// TwinCAT 3 PLC project test
// ProgramVersion: 3.1.4026.27
// libraries:
//   Tc2_Standard, * (Beckhoff Automation GmbH)
//   Tc2_System, * (Beckhoff Automation GmbH)
//   Tc2_Utilities, * (Beckhoff Automation GmbH)
//   Tc3_IotBase, * (Beckhoff Automation GmbH)
//   Tc3_JsonXml, * (Beckhoff Automation GmbH)
//   TcOtlp, * (S&E Engineering)
//   TcUnit, * (www.tcunit.org)
// project tree:
//   / MAIN.TcPOU, PlcTask.TcTTO
//   TEST/TRACING/EXPORTING/ FB_SpanExporter_ForInspection.TcPOU, FB_TestSpanFileExporter.TcPOU, FB_TestSpanSimulation.TcPOU, FB_TestSpanConsoleExporter.TcPOU, FB_TestSpanHttpExporter.TcPOU
//   TEST/EXPORTING/ FB_TestHttpUrlParser.TcPOU
//   TEST/TRACING/TRACESTATE/ FB_TestTraceState.TcPOU
//   TEST/TRACING/PROPAGATION/ FB_TestTraceContextPropagator.TcPOU, FB_TestAdsLoopbackPropagation.TcPOU
//   TEST/TRACING/SAMPLING/ FB_Sampler_ForInspection.TcPOU, FB_TestSamplers.TcPOU
//   TEST/LOGGING/EXPORTING/ FB_TestFileExporter.TcPOU, FB_TestHttpExporter.TcPOU, FB_TestLogExporters.TcPOU
//   TEST/LOGGING/EXPORTING/UTILS/ FB_LogRecordExporter_File_ForSerializationInspection.TcPOU, FB_LogRecordExporter_ForInspection.TcPOU
//   TEST/LOGGING/LOGGER/ FB_TestLogger.TcPOU
//   TEST/LOGGING/LOG_RECORD/ FB_TestLogRecord.TcPOU, FB_TestLogRecordQueue.TcPOU
//   TEST/LOGGING/PROCESSOR/ FB_TestLogProcessors.TcPOU
//   TEST/LOGGING/PROCESSOR/UTILS/ FB_LogRecordProcessor_ConsolePrinter.TcPOU, FB_LogRecordProcessor_ForBatchInspection.TcPOU, FB_LogRecordProcessor_ForRecordInspection.TcPOU, FB_LogRecordProcessor_ForRecordsInspection.TcPOU
//   TEST/LOGGING/PROVIDER/ FB_TestLoggerProvider.TcPOU
//   TEST/LOGGING/SERIALIZATION/ FB_TestProtoJsonSerializer.TcPOU
//   TEST/TRACING/ID_GENERATOR/ FB_TestIdGenerator.TcPOU
//   TEST/TRACING/PROCESSOR/ FB_SpanProcessor_ForInspection.TcPOU, FB_TestSpanProcessors.TcPOU
//   TEST/TRACING/PROVIDER/ FB_TestTracerProvider.TcPOU, FB_TracerProvider_ForInspection.TcPOU
//   TEST/TRACING/TRACER/ FB_MockIdGenerator.TcPOU, FB_TestTracer.TcPOU
//   TEST/TRACING/LINK/ FB_TestLinks.TcPOU
//   TEST/TRACING/SERIALIZATION/ FB_TestSpanProtoJsonSerializer.TcPOU
//   TEST/TRACING/SPAN/ FB_TestSpan.TcPOU, FB_TestSpanContext.TcPOU, FB_TestSpanQueue.TcPOU
//   TEST/VALUES/ FB_TestAttributes.TcPOU, FB_TestOtlpValue.TcPOU
// real-time tasks:
//   TASK PlcTask: cycle T#10ms, priority 20, ADS port 350

CONFIGURATION test
    RESOURCE PLC ON TwinCAT3
        TASK PlcTask(INTERVAL := T#10ms, PRIORITY := 20);
        PROGRAM MAIN WITH PlcTask : MAIN;
    END_RESOURCE
END_CONFIGURATION

// ---- MAIN.TcPOU
PROGRAM MAIN
VAR
	{attribute 'analysis' := '-33'}fbTestOtlpValue: FB_TestOtlpValue();
	{attribute 'analysis' := '-33'}fbTestAttributes: FB_TestAttributes();
	{attribute 'analysis' := '-33'}fbTestLogRecordQueue: FB_TestLogRecordQueue();
	{attribute 'analysis' := '-33'}fbTestLogger: FB_TestLogger();
	{attribute 'analysis' := '-33'}fbTestProvider: FB_TestLoggerProvider();
	{attribute 'analysis' := '-33'}fbTestProcessors: FB_TestLogProcessors();
	{attribute 'analysis' := '-33'}fbTestExporters: FB_TestLogExporters();
	{attribute 'analysis' := '-33'}fbTestLogRecord: FB_TestLogRecord();
	{attribute 'analysis' := '-33'}fbTestProtoJsonSerializer: FB_TestProtoJsonSerializer();
	{attribute 'analysis' := '-33'}fbTestFileExporter: FB_TestFileExporter();
	{attribute 'analysis' := '-33'}fbTestHttpExporter: FB_TestHttpExporter();
	{attribute 'analysis' := '-33'}fbTestIdGenerator: FB_TestIdGenerator();
	{attribute 'analysis' := '-33'}fbTestSpanContext: FB_TestSpanContext();
	{attribute 'analysis' := '-33'}fbTestTraceState: FB_TestTraceState();
	{attribute 'analysis' := '-33'}fbTestTraceContextPropagator: FB_TestTraceContextPropagator();
	{attribute 'analysis' := '-33'}fbTestAdsLoopbackPropagation: FB_TestAdsLoopbackPropagation();
	{attribute 'analysis' := '-33'}fbTestSpan: FB_TestSpan();
	{attribute 'analysis' := '-33'}fbTestTracer: FB_TestTracer();
	{attribute 'analysis' := '-33'}fbTestSpanQueue: FB_TestSpanQueue();
	{attribute 'analysis' := '-33'}fbTestSpanProcessors: FB_TestSpanProcessors();
	{attribute 'analysis' := '-33'}fbTestTracerProvider: FB_TestTracerProvider();
	{attribute 'analysis' := '-33'}fbTestSamplers: FB_TestSamplers();
	{attribute 'analysis' := '-33'}fbTestSpanProtoJsonSerializer: FB_TestSpanProtoJsonSerializer();
	{attribute 'analysis' := '-33'}fbTestLinks: FB_TestLinks();
	{attribute 'analysis' := '-33'}fbTestSpanFileExporter: FB_TestSpanFileExporter();
	{attribute 'analysis' := '-33'}fbTestSpanConsoleExporter: FB_TestSpanConsoleExporter();
	{attribute 'analysis' := '-33'}fbTestSpanHttpExporter: FB_TestSpanHttpExporter();
	{attribute 'analysis' := '-33'}fbTestHttpUrlParser: FB_TestHttpUrlParser();
	{attribute 'analysis' := '-33'}fbTestSpanSimulation: FB_TestSpanSimulation();
END_VAR

TcUnit.RUN();

END_PROGRAM

// ---- TEST/VALUES/FB_TestOtlpValue.TcPOU
(* Tests that ValueFactory validates its inputs, copies what it is given, and that every value it builds is released exactly once. *)
FUNCTION_BLOCK FB_TestOtlpValue EXTENDS FB_TestSuite

THIS^.testCreateStringValidatesInputs();
THIS^.testCreateTraceIdCopiesBytes();
THIS^.testCreateSpanIdCopiesBytes();
THIS^.testCreateKeyValueValidatesInputs();
THIS^.testCreateNumberCopiesEveryNumericType();
THIS^.testCloneCopiesAndForwardsFailures();
THIS^.testDeleteClearsPointer();

(* delete releases a value and clears the caller's pointer, through the concrete or the base type, and refuses a pointer to another value so nothing is released twice. *)
METHOD testDeleteClearsPointer : REFERENCE TO FB_Test
VAR
	pStr: POINTER TO FB_String;
	pOther: POINTER TO FB_String;
	pAny: POINTER TO FB_AnyValue;
	pOtherBefore: POINTER TO FB_String;
	deleted: BOOL;
	failureReason: E_ValueFactoryFailureReason;
END_VAR
TcUnit.TEST('testDeleteClearsPointer');

	// through the concrete pointer type
	IF ValueFactory.createString(pDest:=pStr, pString:=ADR('value'), failureReason=>failureReason) THEN
		deleted := pStr^.delete(pSelf:=pStr);
		THIS^.AssertTrue(deleted, 'Expected delete through an FB_String pointer to succeed');
		THIS^.AssertTrue(pStr = 0, 'Expected delete to clear the FB_String pointer');
	ELSE
		THIS^.AssertTrue(FALSE, 'Expected createString to succeed for the FB_String pointer case');
	END_IF

	// through the abstract base pointer, dispatched to FB_String
	IF ValueFactory.createString(pDest:=pStr, pString:=ADR('value'), failureReason=>failureReason) THEN
		pAny := pStr;
		pStr := 0;
		deleted := pAny^.delete(pSelf:=pAny);
		THIS^.AssertTrue(deleted, 'Expected delete through an FB_AnyValue pointer to succeed');
		THIS^.AssertTrue(pAny = 0, 'Expected delete to clear the FB_AnyValue pointer');
	ELSE
		THIS^.AssertTrue(FALSE, 'Expected createString to succeed for the FB_AnyValue pointer case');
	END_IF

	// a pointer to another value is refused and left untouched
	IF ValueFactory.createString(pDest:=pStr, pString:=ADR('first'), failureReason=>failureReason)
		AND_THEN ValueFactory.createString(pDest:=pOther, pString:=ADR('second'), failureReason=>failureReason)
	THEN
		pOtherBefore := pOther;
		deleted := pStr^.delete(pSelf:=pOther);
		THIS^.AssertFalse(deleted, 'Expected delete with another value$'s pointer to be refused');
		THIS^.AssertTrue(pOther = pOtherBefore, 'Expected a refused delete to leave the pointer unchanged');
		THIS^.AssertEquals_STRING(Expected:='first', Actual:=pStr^.pString^, Message:='Expected the first value to survive a refused delete');
		THIS^.AssertEquals_STRING(Expected:='second', Actual:=pOther^.pString^, Message:='Expected the second value to survive a refused delete');
	ELSE
		THIS^.AssertTrue(FALSE, 'Expected createString to succeed for both strings of the refused delete case');
	END_IF
	IF pStr <> 0 THEN pStr^.delete(pSelf:=pStr); END_IF
	IF pOther <> 0 THEN pOther^.delete(pSelf:=pOther); END_IF

TcUnit.TEST_FINISHED();
END_METHOD

(*
	The clone functions copy strings, numbers, and key values into new allocations.
	A nested clone failure is forwarded with its reason and leaves the destination unassigned, so a caller never gets a half-built value.
*)
METHOD testCloneCopiesAndForwardsFailures : REFERENCE TO FB_Test
VAR
	pStringSource: POINTER TO FB_String;
	pStringClone: POINTER TO FB_String;
	pNumberSource: POINTER TO FB_Number;
	pNumberClone: POINTER TO FB_Number;
	pKeyValueSource: POINTER TO FB_KeyValue;
	pKeyValueClone: POINTER TO FB_KeyValue;
	pAnySource: POINTER TO FB_AnyValue;
	pAnyClone: POINTER TO FB_AnyValue;
	number: DINT := 42;
	success: BOOL;
	failureReason: E_ValueFactoryFailureReason;
	noFailure: E_ValueFactoryFailureReason;
END_VAR
TcUnit.TEST('testCloneCopiesAndForwardsFailures');

	noFailure := E_ValueFactoryFailureReason.NA;

	// cloneString
	success := ValueFactory.createString(pDest:=pStringSource, pString:=ADR('source'), failureReason=>failureReason);
	THIS^.AssertTrue(success AND_THEN failureReason=noFailure AND_THEN pStringSource<>0, 'Expected createString to build the source string');

	success := ValueFactory.cloneString(pDest:=pStringClone, pSrc:=pStringSource, failureReason=>failureReason);
	THIS^.AssertTrue(success AND_THEN failureReason=noFailure AND_THEN pStringClone<>0, 'Expected cloneString to succeed');
	IF pStringClone <> 0 THEN
		THIS^.AssertEquals_STRING('source', pStringClone^.pString^, 'Expected cloneString to copy the source text');
		pStringClone^.delete(pSelf:=pStringClone);
	END_IF

	// cloneNumber
	success := ValueFactory.createNumber(pDest:=pNumberSource, value:=number, failureReason=>failureReason);
	THIS^.AssertTrue(success AND_THEN failureReason=noFailure AND_THEN pNumberSource<>0, 'Expected createNumber to build the source number');

	success := ValueFactory.cloneNumber(pDest:=pNumberClone, pSrc:=pNumberSource, failureReason=>failureReason);
	THIS^.AssertTrue(success AND_THEN failureReason=noFailure AND_THEN pNumberClone<>0, 'Expected cloneNumber to succeed');
	IF pNumberClone <> 0 THEN
		THIS^.AssertTrue(MEMCMP(pNumberClone^.value.pValue, ADR(number), SIZEOF(number))=0, 'Expected cloneNumber to copy the source value');
		pNumberClone^.delete(pSelf:=pNumberClone);
	END_IF

	// cloneAnyValue dispatches on the value type
	pAnySource := pNumberSource;
	success := ValueFactory.cloneAnyValue(pDest:=pAnyClone, pSrc:=pAnySource, failureReason=>failureReason);
	THIS^.AssertTrue(success AND_THEN failureReason=noFailure AND_THEN pAnyClone<>0, 'Expected cloneAnyValue to forward a successful number clone');
	IF pAnyClone <> 0 THEN
		THIS^.AssertTrue(pAnyClone^.eType=E_ValueType.E_Number, 'Expected cloneAnyValue to produce a number');
		pAnyClone^.delete(pSelf:=pAnyClone);
	END_IF

	// cloneKeyValue
	success := ValueFactory.createKeyValue(pDest:=pKeyValueSource, pKey:=ADR('key'), pVal:=pStringSource, failureReason=>failureReason);
	THIS^.AssertTrue(success AND_THEN failureReason=noFailure AND_THEN pKeyValueSource<>0, 'Expected createKeyValue to build the source key value');

	success := ValueFactory.cloneKeyValue(pDest:=pKeyValueClone, pSrc:=pKeyValueSource, failureReason=>failureReason);
	THIS^.AssertTrue(success AND_THEN failureReason=noFailure AND_THEN pKeyValueClone<>0, 'Expected cloneKeyValue to succeed');
	IF pKeyValueClone <> 0 THEN
		THIS^.AssertEquals_STRING('key', pKeyValueClone^.pKey^, 'Expected cloneKeyValue to copy the source key');
		pKeyValueClone^.delete(pSelf:=pKeyValueClone);
	END_IF

	// cloneAnyValue must forward a nested cloneString failure without assigning the destination.
	// free() empties the source string, a state the factory would never build, so the nested clone fails.
	IF pStringSource <> 0 THEN pStringSource^.free(); END_IF
	pAnySource := pStringSource;
	success := ValueFactory.cloneAnyValue(pDest:=pAnyClone, pSrc:=pAnySource, failureReason=>failureReason);
	THIS^.AssertFalse(success, 'Expected cloneAnyValue to reject a string with a null payload');
	THIS^.AssertTrue(failureReason=E_ValueFactoryFailureReason.STRING_POINTER_NULL, 'Expected cloneAnyValue to forward the cloneString failure reason');
	THIS^.AssertTrue(pAnyClone=0, 'Expected a failed cloneAnyValue to leave the destination unassigned');

	// cloneKeyValue must forward the nested createKeyValue failure reason.
	// free() empties the source key value, so it has no key to clone.
	IF pKeyValueSource <> 0 THEN pKeyValueSource^.free(); END_IF
	success := ValueFactory.cloneKeyValue(pDest:=pKeyValueClone, pSrc:=pKeyValueSource, failureReason=>failureReason);
	THIS^.AssertFalse(success, 'Expected cloneKeyValue to reject a key value with a null key');
	THIS^.AssertTrue(failureReason=E_ValueFactoryFailureReason.KEY_POINTER_NULL, 'Expected cloneKeyValue to forward the createKeyValue failure reason');
	THIS^.AssertTrue(pKeyValueClone=0, 'Expected a failed cloneKeyValue to leave the destination unassigned');

	IF pStringSource <> 0 THEN pStringSource^.delete(pSelf:=pStringSource); END_IF
	IF pNumberSource <> 0 THEN pNumberSource^.delete(pSelf:=pNumberSource); END_IF
	IF pKeyValueSource <> 0 THEN pKeyValueSource^.delete(pSelf:=pKeyValueSource); END_IF

TcUnit.TEST_FINISHED();
END_METHOD

(*
	createKeyValue rejects a null key, a null value, or an assigned destination with a distinct reason and allocates nothing.
	On success the key value owns its own copy of the value, so the caller may delete the original.
*)
METHOD testCreateKeyValueValidatesInputs : REFERENCE TO FB_Test
VAR
	pKeyVal: POINTER TO FB_KeyValue;
	pVal: POINTER TO FB_String;
	anyValue: POINTER TO FB_AnyValue;
	expectedType: E_ValueType := E_ValueType.E_KeyValue;
	actualType: E_ValueType;
	pOriginal: POINTER TO FB_KeyValue;
	success: BOOL;
	failureReason: E_ValueFactoryFailureReason;
	noFailure: E_ValueFactoryFailureReason;
	failureCode: INT;
END_VAR
TcUnit.TEST('testCreateKeyValueValidatesInputs');
	noFailure := E_ValueFactoryFailureReason.NA;

	// null key and null value are rejected
	success := ValueFactory.createKeyValue(pDest:=pKeyVal, pKey:=0, pVal:=0, failureReason=>failureReason);
	THIS^.AssertFalse(success, 'Expected createKeyValue to reject a null key pointer');
	THIS^.AssertTrue(failureReason=E_ValueFactoryFailureReason.KEY_POINTER_NULL, 'Expected the null key failure reason');
	THIS^.AssertTrue(pKeyVal=0, 'Expected a null key to leave the destination unassigned');

	success := ValueFactory.createKeyValue(pDest:=pKeyVal, pKey:=ADR('Key'), pVal:=0, failureReason=>failureReason);
	THIS^.AssertFalse(success, 'Expected createKeyValue to reject a null value pointer');
	THIS^.AssertTrue(failureReason=E_ValueFactoryFailureReason.VALUE_POINTER_NULL, 'Expected the null value failure reason');
	THIS^.AssertTrue(pKeyVal=0, 'Expected a null value to leave the destination unassigned');

	// a valid key and value
	success := ValueFactory.createString(pDest:=pVal, pString:=ADR('Value'), failureReason=>failureReason);
	THIS^.AssertTrue(success AND_THEN failureReason=noFailure AND_THEN pVal<>0, 'Expected createString to build the source value');
	success := ValueFactory.createKeyValue(pDest:=pKeyVal, pKey:=ADR('Key'), pVal:=pVal, failureReason=>failureReason);
	THIS^.AssertTrue(success, 'Expected createKeyValue to succeed with a valid key and value');
	THIS^.AssertTrue(failureReason=noFailure, 'Expected a successful createKeyValue to clear the failure reason');
	THIS^.AssertTrue(pKeyVal<>0, 'Expected a successful createKeyValue to allocate the destination');

	// an assigned destination is refused and left as it was
	pOriginal := pKeyVal;
	success := ValueFactory.createKeyValue(pDest:=pKeyVal, pKey:=ADR('Key'), pVal:=pVal, failureReason=>failureReason);
	THIS^.AssertFalse(success, 'Expected createKeyValue to reject an assigned destination');
	THIS^.AssertTrue(failureReason=E_ValueFactoryFailureReason.DESTINATION_ALREADY_ASSIGNED, 'Expected the assigned destination failure reason');
	THIS^.AssertTrue(pKeyVal=pOriginal, 'Expected a refused createKeyValue to keep the existing destination');
	// E_ValueFactoryFailureReason is numbered implicitly after NA := 0; this pins the first failure code at 1
	// so the numeric codes seen in logs and on an HMI do not shift if the enum declaration is edited.
	failureCode := E_ValueFactoryFailureReason.DESTINATION_ALREADY_ASSIGNED;
	THIS^.AssertEquals_INT(1, failureCode, 'Expected the first ValueFactory failure code to be 1');

 	IF pVal <> 0 AND pKeyVal <> 0 THEN
		// a key value is an FB_AnyValue of type E_KeyValue
		anyValue := pKeyVal;
		actualType := anyValue^.eType;
		THIS^.AssertEquals(
			expectedType,
			actualType,
			'Expected the key value to report the E_KeyValue type'
		);
		THIS^.AssertEquals_STRING(
			Actual:=pKeyVal^.pKey^,
			Expected:='Key',
			Message:='Expected the key value to hold the key'
		);
		// deleting the caller's value proves the key value holds its own copy
		pVal^.delete(pSelf:=pVal);
		pVal := pKeyVal^.pVal;
		THIS^.AssertEquals_STRING(
			Actual:=pVal^.pString^,
			Expected:='Value',
			Message:='Expected the key value to keep its value after the original is deleted'
		);
	END_IF
	// cleanup data
	IF pKeyVal <> 0 THEN pKeyVal^.delete(pSelf:=pKeyVal);
	ELSIF pVal <> 0 THEN pVal^.delete(pSelf:=pVal); END_IF


TcUnit.TEST_FINISHED();
END_METHOD

(*
	createNumber accepts every IEC numeric type and keeps its type class and its own copy of the bytes, so the serializer can write the exact type the caller used.
	It also refuses an assigned destination, and free releases the owned data.
*)
METHOD testCreateNumberCopiesEveryNumericType : REFERENCE TO FB_Test
VAR
	nSInt: SINT := -12;
	nInt: INT := -1234;
	nDInt: DINT := -12345;
	nLInt: LINT := -123456;
	nUSInt: USINT := 12;
	nUInt: UINT := 1234;
	nUDInt: UDINT := 12345;
	nULInt: ULINT := 123456;
	fReal: REAL := 42.25;
	fLReal: LREAL := 24.5;
	pValue: POINTER TO FB_Number;
	pDInt: POINTER TO DINT;
	pOriginal: POINTER TO FB_Number;
	anyValue: POINTER TO FB_AnyValue;
	success: BOOL;
	failureReason: E_ValueFactoryFailureReason;
	noFailure: E_ValueFactoryFailureReason;
END_VAR
TcUnit.TEST('testCreateNumberCopiesEveryNumericType');
noFailure := E_ValueFactoryFailureReason.NA;

// ANY_NUM accepts every signed, unsigned, and floating-point IEC numeric type.

// SINT
success := ValueFactory.createNumber(pDest:=pValue, value:=nSInt, failureReason=>failureReason);
THIS^.AssertTrue(success AND_THEN failureReason=noFailure AND_THEN pValue<>0, 'Expected createNumber to accept a SINT');
IF pValue <> 0 THEN
	THIS^.AssertTrue(pValue^.value.typeclass=__SYSTEM.TYPE_CLASS.TYPE_SINT, 'Expected the SINT type to be kept');
	THIS^.AssertTrue(pValue^.value.diSize=SIZEOF(nSInt) AND_THEN MEMCMP(pValue^.value.pValue, ADR(nSInt), SIZEOF(nSInt))=0, 'Expected the SINT value to be copied');
	pValue^.delete(pSelf:=pValue);
END_IF

// INT
success := ValueFactory.createNumber(pDest:=pValue, value:=nInt, failureReason=>failureReason);
THIS^.AssertTrue(success AND_THEN failureReason=noFailure AND_THEN pValue<>0, 'Expected createNumber to accept an INT');
IF pValue <> 0 THEN
	THIS^.AssertTrue(pValue^.value.typeclass=__SYSTEM.TYPE_CLASS.TYPE_INT, 'Expected the INT type to be kept');
	THIS^.AssertTrue(pValue^.value.diSize=SIZEOF(nInt) AND_THEN MEMCMP(pValue^.value.pValue, ADR(nInt), SIZEOF(nInt))=0, 'Expected the INT value to be copied');
	pValue^.delete(pSelf:=pValue);
END_IF

// DINT, plus copy independence and an assigned destination
success := ValueFactory.createNumber(pDest:=pValue, value:=nDInt, failureReason=>failureReason);
THIS^.AssertTrue(success AND_THEN failureReason=noFailure AND_THEN pValue<>0, 'Expected createNumber to accept a DINT');
IF pValue <> 0 THEN
	THIS^.AssertTrue(pValue^.value.typeclass=__SYSTEM.TYPE_CLASS.TYPE_DINT, 'Expected the DINT type to be kept');
	THIS^.AssertTrue(pValue^.value.diSize=SIZEOF(nDInt) AND_THEN MEMCMP(pValue^.value.pValue, ADR(nDInt), SIZEOF(nDInt))=0, 'Expected the DINT value to be copied');
	// The wrapper owns a copy; changing the source must not change the wrapped value.
	pDInt := pValue^.value.pValue;
	nDInt := 7;
	THIS^.AssertEquals_DINT(-12345, pDInt^, 'Expected the number to keep its value after the source DINT changes');
	// A factory call must never replace an already allocated destination.
	pOriginal := pValue;
	success := ValueFactory.createNumber(pDest:=pValue, value:=fLReal, failureReason=>failureReason);
	THIS^.AssertFalse(success, 'Expected createNumber to reject an allocated destination');
	THIS^.AssertTrue(failureReason=E_ValueFactoryFailureReason.DESTINATION_ALREADY_ASSIGNED, 'Expected the assigned number destination failure reason');
	THIS^.AssertTrue(pValue=pOriginal, 'Expected a refused createNumber to keep the existing destination');
	pValue^.delete(pSelf:=pValue);
END_IF

// LINT, which also proves the previous failure reason is cleared
success := ValueFactory.createNumber(pDest:=pValue, value:=nLInt, failureReason=>failureReason);
THIS^.AssertTrue(success AND_THEN failureReason=noFailure AND_THEN pValue<>0, 'Expected createNumber to accept a LINT and clear the previous failure reason');
IF pValue <> 0 THEN
	THIS^.AssertTrue(pValue^.value.typeclass=__SYSTEM.TYPE_CLASS.TYPE_LINT, 'Expected the LINT type to be kept');
	THIS^.AssertTrue(pValue^.value.diSize=SIZEOF(nLInt) AND_THEN MEMCMP(pValue^.value.pValue, ADR(nLInt), SIZEOF(nLInt))=0, 'Expected the LINT value to be copied');
	pValue^.delete(pSelf:=pValue);
END_IF

// USINT
success := ValueFactory.createNumber(pDest:=pValue, value:=nUSInt, failureReason=>failureReason);
THIS^.AssertTrue(success AND_THEN failureReason=noFailure AND_THEN pValue<>0, 'Expected createNumber to accept a USINT');
IF pValue <> 0 THEN
	THIS^.AssertTrue(pValue^.value.typeclass=__SYSTEM.TYPE_CLASS.TYPE_USINT, 'Expected the USINT type to be kept');
	THIS^.AssertTrue(pValue^.value.diSize=SIZEOF(nUSInt) AND_THEN MEMCMP(pValue^.value.pValue, ADR(nUSInt), SIZEOF(nUSInt))=0, 'Expected the USINT value to be copied');
	pValue^.delete(pSelf:=pValue);
END_IF

// UINT
success := ValueFactory.createNumber(pDest:=pValue, value:=nUInt, failureReason=>failureReason);
THIS^.AssertTrue(success AND_THEN failureReason=noFailure AND_THEN pValue<>0, 'Expected createNumber to accept a UINT');
IF pValue <> 0 THEN
	THIS^.AssertTrue(pValue^.value.typeclass=__SYSTEM.TYPE_CLASS.TYPE_UINT, 'Expected the UINT type to be kept');
	THIS^.AssertTrue(pValue^.value.diSize=SIZEOF(nUInt) AND_THEN MEMCMP(pValue^.value.pValue, ADR(nUInt), SIZEOF(nUInt))=0, 'Expected the UINT value to be copied');
	pValue^.delete(pSelf:=pValue);
END_IF

// UDINT
success := ValueFactory.createNumber(pDest:=pValue, value:=nUDInt, failureReason=>failureReason);
THIS^.AssertTrue(success AND_THEN failureReason=noFailure AND_THEN pValue<>0, 'Expected createNumber to accept a UDINT');
IF pValue <> 0 THEN
	THIS^.AssertTrue(pValue^.value.typeclass=__SYSTEM.TYPE_CLASS.TYPE_UDINT, 'Expected the UDINT type to be kept');
	THIS^.AssertTrue(pValue^.value.diSize=SIZEOF(nUDInt) AND_THEN MEMCMP(pValue^.value.pValue, ADR(nUDInt), SIZEOF(nUDInt))=0, 'Expected the UDINT value to be copied');
	pValue^.delete(pSelf:=pValue);
END_IF

// ULINT
success := ValueFactory.createNumber(pDest:=pValue, value:=nULInt, failureReason=>failureReason);
THIS^.AssertTrue(success AND_THEN failureReason=noFailure AND_THEN pValue<>0, 'Expected createNumber to accept a ULINT');
IF pValue <> 0 THEN
	THIS^.AssertTrue(pValue^.value.typeclass=__SYSTEM.TYPE_CLASS.TYPE_ULINT, 'Expected the ULINT type to be kept');
	THIS^.AssertTrue(pValue^.value.diSize=SIZEOF(nULInt) AND_THEN MEMCMP(pValue^.value.pValue, ADR(nULInt), SIZEOF(nULInt))=0, 'Expected the ULINT value to be copied');
	pValue^.delete(pSelf:=pValue);
END_IF

// REAL
success := ValueFactory.createNumber(pDest:=pValue, value:=fReal, failureReason=>failureReason);
THIS^.AssertTrue(success AND_THEN failureReason=noFailure AND_THEN pValue<>0, 'Expected createNumber to accept a REAL');
IF pValue <> 0 THEN
	THIS^.AssertTrue(pValue^.value.typeclass=__SYSTEM.TYPE_CLASS.TYPE_REAL, 'Expected the REAL type to be kept');
	THIS^.AssertTrue(pValue^.value.diSize=SIZEOF(fReal) AND_THEN MEMCMP(pValue^.value.pValue, ADR(fReal), SIZEOF(fReal))=0, 'Expected the REAL value to be copied');
	pValue^.delete(pSelf:=pValue);
END_IF

// LREAL, plus the FB_AnyValue type and free
success := ValueFactory.createNumber(pDest:=pValue, value:=fLReal, failureReason=>failureReason);
THIS^.AssertTrue(success AND_THEN failureReason=noFailure AND_THEN pValue<>0, 'Expected createNumber to accept an LREAL');
IF pValue <> 0 THEN
	THIS^.AssertTrue(pValue^.value.typeclass=__SYSTEM.TYPE_CLASS.TYPE_LREAL, 'Expected the LREAL type to be kept');
	THIS^.AssertTrue(pValue^.value.diSize=SIZEOF(fLReal) AND_THEN MEMCMP(pValue^.value.pValue, ADR(fLReal), SIZEOF(fLReal))=0, 'Expected the LREAL value to be copied');
	// Number values are valid AnyValue instances and participate in the common lifecycle.
	anyValue := pValue;
	THIS^.AssertTrue(anyValue^.eType=E_ValueType.E_Number, 'Expected the number to report the E_Number type');
	anyValue^.free();
	THIS^.AssertTrue(pValue^.value.pValue=0 AND pValue^.value.diSize=0, 'Expected free to clear the owned number data');
	pValue^.delete(pSelf:=pValue);
END_IF

TcUnit.TEST_FINISHED();
END_METHOD

(*
	createSpanId rejects missing or short input and an assigned destination, and otherwise copies the first 8 bytes.
	The span id must hold its own copy so later changes to the caller's buffer cannot alter an emitted id.
*)
METHOD testCreateSpanIdCopiesBytes : REFERENCE TO FB_Test
VAR
	_flag: BOOL;
	_idx: USINT;
	expected: ARRAY [0..spanIdLen-1] OF BYTE;
	pValue: POINTER TO FB_SpanId;
	expectedType: E_ValueType := E_ValueType.E_SpanId;
	actualType: E_ValueType;
	guid_: GUID;
	anyValue: I_OtlpValue;
	pOriginal: POINTER TO FB_SpanId;
	success: BOOL;
	failureReason: E_ValueFactoryFailureReason;
	noFailure: E_ValueFactoryFailureReason;
END_VAR

VAR CONSTANT
	spanIdLen: USINT := 8;  // an OTLP span id is 8 bytes
END_VAR
TcUnit.TEST('testCreateSpanIdCopiesBytes');
	noFailure := E_ValueFactoryFailureReason.NA;

	// null bytes and too few bytes are rejected
	success := ValueFactory.createSpanId(pDest:=pValue, pBytes:=0, nSize:=0, failureReason=>failureReason);
	THIS^.AssertFalse(success, 'Expected createSpanId to reject a null byte pointer');
	THIS^.AssertTrue(failureReason=E_ValueFactoryFailureReason.SPAN_ID_BYTES_POINTER_NULL, 'Expected the null span id byte pointer failure reason');
	THIS^.AssertTrue(pValue=0, 'Expected null span id bytes to leave the destination unassigned');

	success := ValueFactory.createSpanId(pDest:=pValue, pBytes:=ADR(guid_), nSize:=spanIdLen-1, failureReason=>failureReason);
	THIS^.AssertFalse(success, 'Expected createSpanId to reject too few bytes');
	THIS^.AssertTrue(failureReason=E_ValueFactoryFailureReason.SPAN_ID_BYTE_COUNT_TOO_SMALL, 'Expected the span id byte count failure reason');
	THIS^.AssertTrue(pValue=0, 'Expected short span id bytes to leave the destination unassigned');

	// a valid FB_SpanId from the 16 byte GUID; only the first 8 bytes are used
	success := ValueFactory.createSpanId(pDest:=pValue, pBytes:=ADR(guid_), nSize:=SIZEOF(guid_), failureReason=>failureReason);
	THIS^.AssertTrue(success, 'Expected createSpanId to succeed with enough bytes');
	THIS^.AssertTrue(failureReason=noFailure, 'Expected a successful createSpanId to clear the failure reason');
	THIS^.AssertTrue(pValue<>0, 'Expected a successful createSpanId to allocate the destination');

	// an assigned destination is refused and left as it was
	pOriginal := pValue;
	success := ValueFactory.createSpanId(pDest:=pValue, pBytes:=ADR(guid_), nSize:=SIZEOF(guid_), failureReason=>failureReason);
	THIS^.AssertFalse(success, 'Expected createSpanId to reject an assigned destination');
	THIS^.AssertTrue(failureReason=E_ValueFactoryFailureReason.DESTINATION_ALREADY_ASSIGNED, 'Expected the assigned span id destination failure reason');
	THIS^.AssertTrue(pValue=pOriginal, 'Expected a refused createSpanId to keep the existing destination');

 	IF pValue <> 0 THEN
		anyValue := pValue^;
		actualType := anyValue.eType;
		THIS^.AssertEquals(
			expectedType,
			actualType,
			'Expected the span id to report the E_SpanId type'
		);
		MEMCPY(ADR(expected), ADR(guid_), spanIdLen);
		THIS^.AssertEquals(
			expected,
			pValue^.bytes,
			'Expected the span id to hold the source bytes'
		);
		// changing the source GUID must not change the span id, because it holds a copy
		guid_.Data1 := 5;  // changes the first source byte from 0 to 5
		MEMCPY(ADR(expected), ADR(guid_), spanIdLen);
		_flag := TRUE;  // TRUE while every byte still matches the changed source
		FOR _idx := 0 TO spanIdLen-1 DO
			IF pValue^.bytes[_idx] <> expected[_idx] THEN
				_flag := FALSE;
				EXIT;
			END_IF
		END_FOR
		THIS^.AssertFalse(
			_flag,
			'Expected the span id to keep its bytes after the source changes'
		);

		pValue^.delete(pSelf:=pValue);
 END_IF

TcUnit.TEST_FINISHED();
END_METHOD

(* createString rejects a null string or an assigned destination and otherwise copies the text; free then releases the copy. *)
METHOD testCreateStringValidatesInputs : REFERENCE TO FB_Test
VAR
	actual: STRING;
	expected: STRING;
	pValue: POINTER TO FB_String;
	anyValue: POINTER TO FB_AnyValue;
	value: I_OtlpValue;
	pOriginal: POINTER TO FB_String;
	success: BOOL;
	failureReason: E_ValueFactoryFailureReason;
	noFailure: E_ValueFactoryFailureReason;
END_VAR
TcUnit.TEST('testCreateStringValidatesInputs');
	noFailure := E_ValueFactoryFailureReason.NA;

	// a null string is rejected
	success := ValueFactory.createString(pDest:=pValue, pString:=0, failureReason=>failureReason);
	THIS^.AssertFalse(success, 'Expected createString to reject a null string pointer');
	THIS^.AssertTrue(failureReason=E_ValueFactoryFailureReason.STRING_POINTER_NULL, 'Expected the null string failure reason');
	THIS^.AssertTrue(pValue=0, 'Expected a null string to leave the destination unassigned');

	// a valid FB_String
	success := ValueFactory.createString(pDest:=pValue, pString:=ADR('FB_String'), failureReason=>failureReason);
	THIS^.AssertTrue(success, 'Expected createString to succeed with a valid string');
	THIS^.AssertTrue(failureReason=noFailure, 'Expected a successful createString to clear the previous failure reason');
	THIS^.AssertTrue(pValue<>0, 'Expected a successful createString to allocate the destination');

	// an assigned destination is refused and left as it was
	pOriginal := pValue;
	success := ValueFactory.createString(pDest:=pValue, pString:=ADR('FB_String'), failureReason=>failureReason);
	THIS^.AssertFalse(success, 'Expected createString to reject an assigned destination');
	THIS^.AssertTrue(failureReason=E_ValueFactoryFailureReason.DESTINATION_ALREADY_ASSIGNED, 'Expected the assigned string destination failure reason');
	THIS^.AssertTrue(pValue=pOriginal, 'Expected a refused createString to keep the existing destination');

	// the string holds the copied text
	THIS^.AssertTrue(pValue <> 0, 'Expected the string to still be allocated after the refused create');
	IF pValue <> 0 THEN
		// the value can be used as an FB_AnyValue and an I_OtlpValue
		anyValue := pValue;
		value := pValue^;
		actual := pValue^.pString^;
		expected := 'FB_String';
		THIS^.AssertEquals(
			expected,
			actual,
			'Expected the string to hold the copied text'
		);
		// free through the interface releases the owned text
		value.free();
		THIS^.AssertTrue(pValue^.pString = 0, 'Expected free to clear the string pointer');
		pValue^.delete(pSelf:=pValue);
 END_IF

TcUnit.TEST_FINISHED();
END_METHOD

(*
	createTraceId rejects missing or short input and an assigned destination, and otherwise copies 16 bytes.
	The trace id must hold its own copy so later changes to the caller's buffer cannot alter an emitted id.
*)
METHOD testCreateTraceIdCopiesBytes : REFERENCE TO FB_Test
VAR
	_flag: BOOL;
	_idx: USINT;
	expected: ARRAY [0..traceIdLen-1] OF BYTE;
	expectedType: E_ValueType := E_ValueType.E_TraceId;
	actualType: E_ValueType;
	pValue: POINTER TO FB_TraceId;
	guid_: GUID;
	anyValue: I_OtlpValue;
	pOriginal: POINTER TO FB_TraceId;
	success: BOOL;
	failureReason: E_ValueFactoryFailureReason;
	noFailure: E_ValueFactoryFailureReason;
END_VAR

VAR CONSTANT
	traceIdLen: USINT := 16;  // an OTLP trace id is 16 bytes
END_VAR
TcUnit.TEST('testCreateTraceIdCopiesBytes');
	noFailure := E_ValueFactoryFailureReason.NA;
	// null bytes and too few bytes are rejected
	success := ValueFactory.createTraceId(pDest:=pValue, pBytes:=0, nSize:=0, failureReason=>failureReason);
	THIS^.AssertFalse(success, 'Expected createTraceId to reject a null byte pointer');
	THIS^.AssertTrue(failureReason=E_ValueFactoryFailureReason.TRACE_ID_BYTES_POINTER_NULL, 'Expected the null trace id byte pointer failure reason');
	THIS^.AssertTrue(pValue=0, 'Expected null trace id bytes to leave the destination unassigned');

	success := ValueFactory.createTraceId(pDest:=pValue, pBytes:=ADR(guid_), nSize:=traceIdLen-1, failureReason=>failureReason);
	THIS^.AssertFalse(success, 'Expected createTraceId to reject too few bytes');
	THIS^.AssertTrue(failureReason=E_ValueFactoryFailureReason.TRACE_ID_BYTE_COUNT_TOO_SMALL, 'Expected the trace id byte count failure reason');
	THIS^.AssertTrue(pValue=0, 'Expected short trace id bytes to leave the destination unassigned');

	// a valid FB_TraceId from the 16 byte GUID
	success := ValueFactory.createTraceId(pDest:=pValue, pBytes:=ADR(guid_), nSize:=SIZEOF(guid_), failureReason=>failureReason);
	THIS^.AssertTrue(success, 'Expected createTraceId to succeed with enough bytes');
	THIS^.AssertTrue(failureReason=noFailure, 'Expected a successful createTraceId to clear the failure reason');
	THIS^.AssertTrue(pValue<>0, 'Expected a successful createTraceId to allocate the destination');

	// an assigned destination is refused and left as it was
	pOriginal := pValue;
	success := ValueFactory.createTraceId(pDest:=pValue, pBytes:=ADR(guid_), nSize:=SIZEOF(guid_), failureReason=>failureReason);
	THIS^.AssertFalse(success, 'Expected createTraceId to reject an assigned destination');
	THIS^.AssertTrue(failureReason=E_ValueFactoryFailureReason.DESTINATION_ALREADY_ASSIGNED, 'Expected the assigned trace id destination failure reason');
	THIS^.AssertTrue(pValue=pOriginal, 'Expected a refused createTraceId to keep the existing destination');

 	IF pValue <> 0 THEN
		// the trace id can be used as an I_OtlpValue
		anyValue := pValue^;
		actualType := anyValue.eType;
		THIS^.AssertEquals(
			expectedType,
			actualType,
			'Expected the trace id to report the E_TraceId type'
		);
		MEMCPY(ADR(expected), ADR(guid_), traceIdLen);
		THIS^.AssertEquals(
			expected,
			pValue^.bytes,
			'Expected the trace id to hold the source bytes'
		);
		// changing the source GUID must not change the trace id, because it holds a copy
		guid_.Data1 := 5;  // changes the first source byte from 0 to 5
		MEMCPY(ADR(expected), ADR(guid_), traceIdLen);
		_flag := TRUE;  // TRUE while every byte still matches the changed source
		FOR _idx := 0 TO traceIdLen-1 DO
			IF pValue^.bytes[_idx] <> expected[_idx] THEN
				_flag := FALSE;
				EXIT;
			END_IF
		END_FOR
		THIS^.AssertFalse(
			_flag,
			'Expected the trace id to keep its bytes after the source changes'
		);
		pValue^.free();
		pValue^.delete(pSelf:=pValue);
 END_IF

TcUnit.TEST_FINISHED();
END_METHOD

END_FUNCTION_BLOCK

// ---- TEST/VALUES/FB_TestAttributes.TcPOU
(* Tests attribute value creation, ownership, and copying. *)
FUNCTION_BLOCK FB_TestAttributes EXTENDS FB_TestSuite

THIS^.testCopyFromIsIndependent();
THIS^.testRejectsInvalidAndExcessAttributes();
THIS^.testGetAttributeBorrowsByKey();
THIS^.testCopyAttributeRenamesAndReplaces();
THIS^.testCopyAttributeRespectsCountLimit();

(*
	copyAttribute into a full collection drops a new key the same way setAttribute does, leaving the
	collection unchanged apart from droppedCount, and still replaces a key the collection already holds.
*)
METHOD testCopyAttributeRespectsCountLimit : REFERENCE TO FB_Test
VAR
	span: FB_Attributes(maxCount:=TcOtlp_GVL.DEFAULT_MAX_ATTRIBUTE_COUNT);
	resource: FB_Attributes(maxCount:=1);
	pKv: POINTER TO FB_KeyValue;
	pStr: POINTER TO FB_String;
	success: BOOL;
	failureReason: E_AttributesFailureReason;
END_VAR
TcUnit.TEST('testCopyAttributeRespectsCountLimit');
	success := span.setStringAttribute(key:='peer.name', value:='modbus-device', failureReason=>failureReason);
	THIS^.AssertTrue(success, 'Expected the source attribute to be added');
	success := resource.setStringAttribute(key:='service.name', value:='PLC1', failureReason=>failureReason);
	THIS^.AssertTrue(success, 'Expected the target attribute to fill the collection');

	// a new key is dropped: the copy is released and only droppedCount changes
	success := resource.copyAttribute(src:=span, key:='peer.name', failureReason=>failureReason);
	THIS^.AssertFalse(success, 'Expected a copy under a new key to be rejected by a full collection');
	THIS^.AssertTrue(failureReason=E_AttributesFailureReason.ATTRIBUTE_COUNT_LIMIT_REACHED, 'Expected the attribute count failure reason');
	THIS^.AssertEquals_UDINT(1, resource.count, 'Expected the rejected copy not to change the count');
	THIS^.AssertEquals_UDINT(1, resource.droppedCount, 'Expected the rejected copy to increment the dropped count');
	THIS^.AssertTrue(resource.getAttribute('peer.name') = 0, 'Expected the rejected key not to be added');
	pKv := resource.getAttribute('service.name');
	IF pKv <> 0 THEN
		pStr := pKv^.pVal;
		THIS^.AssertEquals_STRING('PLC1', pStr^.pString^, 'Expected the rejected copy to leave service.name untouched');
	ELSE
		THIS^.AssertTrue(FALSE, 'Expected service.name to survive the rejected copy');
	END_IF

	// replacing a key the full collection already holds still succeeds
	success := resource.copyAttribute(src:=span, key:='peer.name', destKey:='service.name', failureReason=>failureReason);
	THIS^.AssertTrue(success AND_THEN failureReason=E_AttributesFailureReason.NA, 'Expected a copy onto an existing key to succeed at the limit');
	THIS^.AssertEquals_UDINT(1, resource.count, 'Expected the replacement not to change the count');
	THIS^.AssertEquals_UDINT(1, resource.droppedCount, 'Expected the replacement not to increment the dropped count');
	pKv := resource.getAttribute('service.name');
	IF pKv <> 0 THEN
		pStr := pKv^.pVal;
		THIS^.AssertEquals_STRING('modbus-device', pStr^.pString^, 'Expected service.name to hold the copied value');
	ELSE
		THIS^.AssertTrue(FALSE, 'Expected service.name to exist after the replacement');
	END_IF

	span.free();
	resource.free();
TcUnit.TEST_FINISHED();
END_METHOD

(*
	copyAttribute copies one attribute, under a new name when destKey is given, replacing any
	attribute already held under that name. The copy is independent of the source, and a key the
	source lacks is reported without touching the target.
*)
METHOD testCopyAttributeRenamesAndReplaces : REFERENCE TO FB_Test
VAR
	span: FB_Attributes(maxCount:=TcOtlp_GVL.DEFAULT_MAX_ATTRIBUTE_COUNT);
	resource: FB_Attributes(maxCount:=TcOtlp_GVL.DEFAULT_MAX_ATTRIBUTE_COUNT);
	pKv: POINTER TO FB_KeyValue;
	pStr: POINTER TO FB_String;
	success: BOOL;
	failureReason: E_AttributesFailureReason;
	noFailure: E_AttributesFailureReason;
END_VAR
TcUnit.TEST('testCopyAttributeRenamesAndReplaces');
	noFailure := E_AttributesFailureReason.NA;

	success := span.setStringAttribute(key:='peer.name', value:='modbus-device', failureReason=>failureReason);
	THIS^.AssertTrue(success, 'Expected the source attribute to be added');
	success := resource.setStringAttribute(key:='service.name', value:='PLC1', failureReason=>failureReason);
	THIS^.AssertTrue(success, 'Expected the target attribute to be added');

	// copying under a new name replaces the existing value instead of adding a key
	success := resource.copyAttribute(src:=span, key:='peer.name', destKey:='service.name', failureReason=>failureReason);
	THIS^.AssertTrue(success AND_THEN failureReason=noFailure, 'Expected the renamed copy to succeed');
	THIS^.AssertEquals_UDINT(1, resource.count, 'Expected the renamed copy to replace service.name rather than add a key');
	THIS^.AssertTrue(resource.getAttribute('peer.name') = 0, 'Expected the renamed copy not to add the source key');
	pKv := resource.getAttribute('service.name');
	IF pKv <> 0 THEN
		pStr := pKv^.pVal;
		THIS^.AssertEquals_STRING('modbus-device', pStr^.pString^, 'Expected service.name to hold the copied peer.name value');
	ELSE
		THIS^.AssertTrue(FALSE, 'Expected service.name to exist after the copy');
	END_IF

	// without destKey the attribute keeps its name
	success := resource.copyAttribute(src:=span, key:='peer.name', failureReason=>failureReason);
	THIS^.AssertTrue(success AND_THEN failureReason=noFailure, 'Expected a copy under the same key to succeed');
	THIS^.AssertEquals_UDINT(2, resource.count, 'Expected the copy to add peer.name');
	THIS^.AssertTrue(resource.getAttribute('peer.name') <> 0, 'Expected peer.name in the target');

	// the source is unchanged and freeing it leaves the copies intact
	THIS^.AssertEquals_UDINT(1, span.count, 'Expected copyAttribute to leave the source unchanged');
	span.free();
	pKv := resource.getAttribute('service.name');
	IF pKv <> 0 THEN
		pStr := pKv^.pVal;
		THIS^.AssertEquals_STRING('modbus-device', pStr^.pString^, 'Expected the copy to outlive the freed source');
	ELSE
		THIS^.AssertTrue(FALSE, 'Expected service.name to survive freeing the source');
	END_IF

	// KEY_NOT_FOUND: the source has no such key, and the target is untouched
	success := resource.copyAttribute(src:=span, key:='peer.name', destKey:='service.name', failureReason=>failureReason);
	THIS^.AssertFalse(success, 'Expected a missing source key to be rejected');
	THIS^.AssertTrue(failureReason=E_AttributesFailureReason.KEY_NOT_FOUND, 'Expected the key not found failure reason');
	THIS^.AssertEquals_UDINT(2, resource.count, 'Expected a missing source key not to change the target');

	// a collection can copy one of its own attributes to a new name
	success := resource.copyAttribute(src:=resource, key:='service.name', destKey:='service.alias', failureReason=>failureReason);
	THIS^.AssertTrue(success AND_THEN failureReason=noFailure, 'Expected an in-place copy to succeed');
	THIS^.AssertEquals_UDINT(3, resource.count, 'Expected the in-place copy to add service.alias');

	resource.free();
TcUnit.TEST_FINISHED();
END_METHOD

(* getAttribute finds an attribute by key without taking ownership or moving the next cursor, and returns 0 for a missing key. *)
METHOD testGetAttributeBorrowsByKey : REFERENCE TO FB_Test
VAR
	attributes: FB_Attributes(maxCount:=TcOtlp_GVL.DEFAULT_MAX_ATTRIBUTE_COUNT);
	pKv: POINTER TO FB_KeyValue;
	numVal: REAL := 2;
	success: BOOL;
	failureReason: E_AttributesFailureReason;
END_VAR
TcUnit.TEST('testGetAttributeBorrowsByKey');
	THIS^.AssertTrue(attributes.getAttribute('missing') = 0, 'Expected an empty collection to return 0');

	success := attributes.setStringAttribute(key:='first', value:='one', failureReason=>failureReason);
	THIS^.AssertTrue(success, 'Expected the first attribute to be added');
	success := attributes.setNumberAttribute(key:='second', value:=numVal, failureReason=>failureReason);
	THIS^.AssertTrue(success, 'Expected the second attribute to be added');

	attributes.reset();
	pKv := attributes.getAttribute('second');
	THIS^.AssertTrue(pKv <> 0, 'Expected the second attribute to be found');
	IF pKv <> 0 THEN
		THIS^.AssertEquals_STRING('second', pKv^.pKey^, 'Expected the attribute with the requested key');
	END_IF
	THIS^.AssertTrue(attributes.getAttribute('missing') = 0, 'Expected a missing key to return 0');

	// the cursor has not moved, so next still starts at the first attribute
	pKv := attributes.next();
	IF pKv <> 0 THEN
		THIS^.AssertEquals_STRING('first', pKv^.pKey^, 'Expected getAttribute not to move the next cursor');
	ELSE
		THIS^.AssertTrue(FALSE, 'Expected next to return the first attribute');
	END_IF
	THIS^.AssertEquals_UDINT(2, attributes.count, 'Expected getAttribute not to change the collection');

	attributes.free();
TcUnit.TEST_FINISHED();
END_METHOD

(* copyFrom gives the target its own copy of every attribute, so freeing either collection leaves the other intact. *)
METHOD testCopyFromIsIndependent : REFERENCE TO FB_Test
VAR
	attributes: FB_Attributes(maxCount:=TcOtlp_GVL.DEFAULT_MAX_ATTRIBUTE_COUNT);
	copyTarget: FB_Attributes(maxCount:=TcOtlp_GVL.DEFAULT_MAX_ATTRIBUTE_COUNT);
	strVal: T_MaxString := 'String';
	numVal: REAL := 42;
	success: BOOL;
	failureReason: E_AttributesFailureReason;
	noFailure: E_AttributesFailureReason;
END_VAR
TcUnit.TEST('testCopyFromIsIndependent');
	noFailure := E_AttributesFailureReason.NA;

	// adding to the source does not touch the target
	success := attributes.setStringAttribute(key:='strKey', value:=strVal, failureReason=>failureReason);
	THIS^.AssertTrue(success AND_THEN failureReason=noFailure, 'Expected string attribute creation to succeed');
	THIS^.AssertTrue(attributes.count = 1, 'Expected the source to hold one attribute after the string is added');
	THIS^.AssertTrue(copyTarget.count = 0, 'Expected the target to stay empty after the string is added to the source');

	success := attributes.setNumberAttribute(key:='numKey', value:=numVal, failureReason=>failureReason);
	THIS^.AssertTrue(success AND_THEN failureReason=noFailure, 'Expected number attribute creation to succeed');
	THIS^.AssertTrue(attributes.count = 2, 'Expected the source to hold two attributes after the number is added');
	THIS^.AssertTrue(copyTarget.count = 0, 'Expected the target to stay empty after the number is added to the source');

	// copyFrom copies both attributes and leaves the source unchanged
	success := copyTarget.copyFrom(src:=attributes, failureReason=>failureReason);
	THIS^.AssertTrue(success AND_THEN failureReason=noFailure, 'Expected attribute copy to succeed');
	THIS^.AssertTrue(attributes.count = 2, 'Expected copyFrom to leave both attributes in the source');
	THIS^.AssertTrue(copyTarget.count = 2, 'Expected copyFrom to copy both attributes into the target');

	// freeing the source proves the target owns its own copies
	attributes.free();
	THIS^.AssertTrue(attributes.count = 0, 'Expected free to empty the source');
	THIS^.AssertTrue(copyTarget.count = 2, 'Expected the target to keep both attributes after the source is freed');

	copyTarget.free();
	THIS^.AssertTrue(copyTarget.count = 0, 'Expected free to empty the target');
TcUnit.TEST_FINISHED();
END_METHOD

(*
	Each invalid key-value pair, invalid number, and attribute beyond maxCount is rejected with its own failure reason.
	The count limit drops new keys but still lets an existing key be replaced, which bounds memory without losing updates.
*)
METHOD testRejectsInvalidAndExcessAttributes : REFERENCE TO FB_Test
VAR
	attributes: FB_Attributes(maxCount:=1);
	copySource: FB_Attributes(maxCount:=2);
	limitedCopyTarget: FB_Attributes(maxCount:=1);
	invalidKv: FB_KeyValue(pKey:=0, pVal:=0);  // built by hand because ValueFactory refuses a null key or value
	pKv: POINTER TO FB_KeyValue;
	pKey: POINTER TO STRING;
	key: T_MaxString := 'key';
	keySize: UDINT;
	invalidValue: AnyType;
	success: BOOL;
	failureReason: E_AttributesFailureReason;
	noFailure: E_AttributesFailureReason;
	failureCode: UDINT;
END_VAR
TcUnit.TEST('testRejectsInvalidAndExcessAttributes');
	noFailure := E_AttributesFailureReason.NA;

	// KV_POINTER_NULL: no key-value pair at all
	success := attributes.setAttribute(pValue:=pKv, failureReason=>failureReason);
	THIS^.AssertFalse(success, 'Expected a null key-value pointer to be rejected');
	THIS^.AssertTrue(failureReason=E_AttributesFailureReason.KV_POINTER_NULL, 'Expected the null key-value failure reason');

	// KV_KEY_POINTER_NULL: a pair with no key
	pKv := ADR(invalidKv);
	success := attributes.setAttribute(pValue:=pKv, failureReason=>failureReason);
	THIS^.AssertFalse(success, 'Expected a key-value pair without a key to be rejected');
	THIS^.AssertTrue(failureReason=E_AttributesFailureReason.KV_KEY_POINTER_NULL, 'Expected the missing key failure reason');

	// KV_VALUE_POINTER_NULL: a pair with a key but no value
	pKv := 0;
	keySize := LEN2(ADR(key)) + 1;  // + 1 for the null terminator
	pKey := __NEW(BYTE, keySize);
	IF pKey <> 0 THEN
		MEMCPY(pKey, ADR(key), keySize);
		pKv := __NEW(FB_KeyValue(pKey:=pKey, pVal:=0));  // built by hand because ValueFactory refuses a null key or value
		IF pKv <> 0 THEN
			pKey := 0;  // the key-value pair now owns the key
			success := attributes.setAttribute(pValue:=pKv, failureReason=>failureReason);
			THIS^.AssertFalse(success, 'Expected a key-value pair without a value to be rejected');
			THIS^.AssertTrue(failureReason=E_AttributesFailureReason.KV_VALUE_POINTER_NULL, 'Expected the missing value failure reason');
			pKv^.delete(pSelf:=pKv);
		ELSE
			THIS^.AssertTrue(FALSE, 'Expected allocation of the invalid key-value test fixture to succeed');
			__DELETE(pKey);
		END_IF
	ELSE
		THIS^.AssertTrue(FALSE, 'Expected allocation of the invalid key test fixture to succeed');
	END_IF

	// KV_VALUE_INVALID: an empty AnyType carries no number
	success := attributes.setNumberAttribute_AnyType(key:='invalid', value:=invalidValue, failureReason=>failureReason);
	THIS^.AssertFalse(success, 'Expected invalid number data to be rejected');
	THIS^.AssertTrue(failureReason=E_AttributesFailureReason.KV_VALUE_INVALID, 'Expected the invalid value failure reason');

	// ATTRIBUTE_COUNT_LIMIT_REACHED: a new key beyond maxCount (1) is dropped
	success := attributes.setStringAttribute(key:='first', value:='one', failureReason=>failureReason);
	THIS^.AssertTrue(success AND_THEN failureReason=noFailure, 'Expected the first attribute to be added');
	success := attributes.setStringAttribute(key:='second', value:='two', failureReason=>failureReason);
	THIS^.AssertFalse(success, 'Expected the attribute count limit to reject a new key');
	THIS^.AssertTrue(failureReason=E_AttributesFailureReason.ATTRIBUTE_COUNT_LIMIT_REACHED, 'Expected the attribute count failure reason');
	THIS^.AssertEquals_UDINT(1, attributes.count, 'Expected the rejected attribute not to change the count');
	THIS^.AssertEquals_UDINT(1, attributes.droppedCount, 'Expected the rejected attribute to increment the dropped count');

	// replacing an existing key is still allowed at the limit
	success := attributes.setStringAttribute(key:='first', value:='replacement', failureReason=>failureReason);
	THIS^.AssertTrue(success, 'Expected an existing key to be replaceable at the count limit');
	THIS^.AssertTrue(failureReason=noFailure, 'Expected success to clear the prior failure reason');
	THIS^.AssertEquals_UDINT(1, attributes.count, 'Expected replacement not to change the attribute count');
	THIS^.AssertEquals_UDINT(1, attributes.droppedCount, 'Expected replacement not to increment the dropped count');

	// ATTRIBUTE_COUNT_LIMIT_REACHED from copyFrom: two source attributes into a target of maxCount 1
	success := copySource.setStringAttribute(key:='first', value:='one', failureReason=>failureReason);
	THIS^.AssertTrue(success, 'Expected the first source attribute to be added');
	success := copySource.setStringAttribute(key:='second', value:='two', failureReason=>failureReason);
	THIS^.AssertTrue(success, 'Expected the second source attribute to be added');
	success := limitedCopyTarget.copyFrom(src:=copySource, failureReason=>failureReason);
	THIS^.AssertFalse(success, 'Expected copyFrom to reject attributes beyond the destination limit');
	THIS^.AssertTrue(failureReason=E_AttributesFailureReason.ATTRIBUTE_COUNT_LIMIT_REACHED, 'Expected copyFrom to expose the count limit failure reason');
	THIS^.AssertEquals_UDINT(1, limitedCopyTarget.count, 'Expected copyFrom to retain only the attribute copied before failure');

	// E_AttributesFailureReason is numbered implicitly after NA := 0; this pins the first failure code at 1
	// so the numeric codes seen in logs and on an HMI do not shift if the enum declaration is edited.
	failureCode := E_AttributesFailureReason.KV_POINTER_NULL;
	THIS^.AssertEquals_UDINT(1, failureCode, 'Expected the first attributes failure code to be 1');

	attributes.free();
	copySource.free();
	limitedCopyTarget.free();
TcUnit.TEST_FINISHED();
END_METHOD

END_FUNCTION_BLOCK

// ---- TEST/LOGGING/LOG_RECORD/FB_TestLogRecordQueue.TcPOU
(* Tests log record queue behavior and ownership transfer. *)
FUNCTION_BLOCK FB_TestLogRecordQueue EXTENDS FB_TestSuite

THIS^.testEnforcesMaximumSize();
THIS^.testAllowsUnboundedLength();
THIS^.testDropsOldestRecordFirst();
THIS^.testPushAndPopTransferRecordOwnership();
THIS^.testTransfersQueueOwnership();
THIS^.testTransfersRequestedCount();
THIS^.testReportsFailureReasons();

(* A queue built with maxCount 0 is unbounded and accepts every record without dropping; batch processors rely on this when no limit is configured. *)
METHOD testAllowsUnboundedLength : REFERENCE TO FB_Test
VAR
	queue: FB_LogRecordQueue(maxCount:=0);
	pRecord: POINTER TO FB_LogRecord;
	failureReason: E_LogRecordQueueFailureReason;
	success: BOOL;
	_idx: UDINT;
END_VAR
TcUnit.TEST('testAllowsUnboundedLength');
	FOR _idx := 1 TO 3 DO
		// opaque queue node: no factory hands a test an owned FB_LogRecord
		pRecord := __NEW(FB_LogRecord(severityNumber:=E_SeverityNumber.INFO, timestamp:=_idx));
		success := queue.push(pValue:=pRecord, failureReason=>failureReason);
		THIS^.AssertTrue(success AND_THEN pRecord = 0, 'Expected the unbounded queue to take ownership');
	END_FOR
	THIS^.AssertEquals_UDINT(3, queue.count, 'Expected maxSize zero to allow every record');
	THIS^.AssertEquals_UDINT(0, queue.droppedCount, 'Expected the unbounded queue not to drop records');
	queue.free();
TcUnit.TEST_FINISHED();
END_METHOD

(* A full queue drops its oldest record to make room for a new one, so the most recent logs survive a burst. *)
METHOD testDropsOldestRecordFirst : REFERENCE TO FB_Test
VAR
	queue: FB_LogRecordQueue(maxCount:=2);
	pRecord: POINTER TO FB_LogRecord;
	failureReason: E_LogRecordQueueFailureReason;
	success: BOOL;
	_idx: UDINT;
END_VAR
TcUnit.TEST('testDropsOldestRecordFirst');
	FOR _idx := 1 TO 3 DO
		// opaque queue node: no factory hands a test an owned FB_LogRecord
		pRecord := __NEW(FB_LogRecord(severityNumber:=E_SeverityNumber.INFO, timestamp:=_idx));
		success := queue.push(pValue:=pRecord, failureReason=>failureReason);
		THIS^.AssertTrue(success, 'Expected push to succeed');
	END_FOR

	success := queue.pop(pValue:=pRecord, failureReason=>failureReason);
	THIS^.AssertTrue(success AND_THEN pRecord <> 0 AND_THEN pRecord^.timestamp = 2, 'Expected timestamp 1 to be dropped first');
	IF pRecord <> 0 THEN pRecord^.delete(pSelf:=pRecord); END_IF
	success := queue.pop(pValue:=pRecord, failureReason=>failureReason);
	THIS^.AssertTrue(success AND_THEN pRecord <> 0 AND_THEN pRecord^.timestamp = 3, 'Expected the newest record to remain at the tail');
	IF pRecord <> 0 THEN pRecord^.delete(pSelf:=pRecord); END_IF
TcUnit.TEST_FINISHED();
END_METHOD

(* A bounded queue never holds more than maxCount records and counts each record it drops, so memory stays bounded on the PLC. *)
METHOD testEnforcesMaximumSize : REFERENCE TO FB_Test
VAR
	queue: FB_LogRecordQueue(maxCount:=2);
	pRecord: POINTER TO FB_LogRecord;
	failureReason: E_LogRecordQueueFailureReason;
	success: BOOL;
	_idx: UDINT;
END_VAR
TcUnit.TEST('testEnforcesMaximumSize');
	FOR _idx := 1 TO 3 DO
		// opaque queue node: no factory hands a test an owned FB_LogRecord
		pRecord := __NEW(FB_LogRecord(severityNumber:=E_SeverityNumber.INFO, timestamp:=_idx));
		success := queue.push(pValue:=pRecord, failureReason=>failureReason);
		THIS^.AssertTrue(success AND_THEN pRecord = 0, 'Expected push to take ownership');
		THIS^.AssertTrue(queue.count <= queue.maxCount, 'Expected count not to exceed maxSize');
	END_FOR
	THIS^.AssertTrue(queue.count = 2, 'Expected the queue to remain at its maximum size');
	THIS^.AssertTrue(queue.droppedCount = 1, 'Expected one record to be dropped');
TcUnit.TEST_FINISHED();
END_METHOD

(* Push takes ownership of the record and clears the caller's pointer, and pop hands the same record back; each record then has exactly one owner. *)
METHOD testPushAndPopTransferRecordOwnership : REFERENCE TO FB_Test
VAR
	queue: FB_LogRecordQueue(maxCount:=2);
	pRecord: POINTER TO FB_LogRecord;
	pOriginal: POINTER TO FB_LogRecord;
	failureReason: E_LogRecordQueueFailureReason;
	noFailure: E_LogRecordQueueFailureReason;
	success: BOOL;
END_VAR
TcUnit.TEST('testPushAndPopTransferRecordOwnership');
	noFailure := E_LogRecordQueueFailureReason.NA;
	// opaque queue node: no factory hands a test an owned FB_LogRecord
	pRecord := __NEW(FB_LogRecord(severityNumber:=E_SeverityNumber.INFO, timestamp:=42));
	pOriginal := pRecord;
	success := queue.push(pValue:=pRecord, failureReason=>failureReason);
	THIS^.AssertTrue(success AND_THEN failureReason = noFailure, 'Expected push to succeed without a failure reason');
	THIS^.AssertTrue(pRecord = 0 AND_THEN queue.count = 1, 'Expected push to transfer ownership into the queue');

	success := queue.pop(pValue:=pRecord, failureReason=>failureReason);
	THIS^.AssertTrue(success AND_THEN failureReason = noFailure, 'Expected pop to succeed without a failure reason');
	THIS^.AssertTrue(pRecord = pOriginal AND_THEN queue.count = 0, 'Expected pop to transfer the same record back to the caller');
	IF pRecord <> 0 THEN pRecord^.delete(pSelf:=pRecord); END_IF
TcUnit.TEST_FINISHED();
END_METHOD

(* Push and pop refuse a null record, an empty queue and an already assigned destination with a distinct reason each, and a later success clears the reason. *)
METHOD testReportsFailureReasons : REFERENCE TO FB_Test
VAR
	queue: FB_LogRecordQueue(maxCount:=1);
	pRecord: POINTER TO FB_LogRecord;
	pAssigned: POINTER TO FB_LogRecord;
	failureReason: E_LogRecordQueueFailureReason;
	noFailure: E_LogRecordQueueFailureReason;
	success: BOOL;
END_VAR
TcUnit.TEST('testReportsFailureReasons');
	noFailure := E_LogRecordQueueFailureReason.NA;
	success := queue.push(pValue:=pRecord, failureReason=>failureReason);
	THIS^.AssertFalse(success, 'Expected a null record push to fail');
	THIS^.AssertTrue(failureReason = E_LogRecordQueueFailureReason.RECORD_POINTER_NULL, 'Expected the null record failure reason');

	success := queue.pop(pValue:=pRecord, failureReason=>failureReason);
	THIS^.AssertFalse(success, 'Expected an empty pop to fail');
	THIS^.AssertTrue(failureReason = E_LogRecordQueueFailureReason.QUEUE_EMPTY, 'Expected the empty queue failure reason');

	// opaque queue node: no factory hands a test an owned FB_LogRecord
	pAssigned := __NEW(FB_LogRecord(severityNumber:=E_SeverityNumber.INFO, timestamp:=2));
	success := queue.pop(pValue:=pAssigned, failureReason=>failureReason);
	THIS^.AssertFalse(success, 'Expected pop into an assigned pointer to fail');
	THIS^.AssertTrue(failureReason = E_LogRecordQueueFailureReason.DESTINATION_ALREADY_ASSIGNED, 'Expected the assigned destination failure reason');
	IF pAssigned <> 0 THEN pAssigned^.delete(pSelf:=pAssigned); END_IF

	pRecord := __NEW(FB_LogRecord(severityNumber:=E_SeverityNumber.INFO, timestamp:=5));
	success := queue.push(pValue:=pRecord, failureReason=>failureReason);
	THIS^.AssertTrue(success AND_THEN failureReason = noFailure, 'Expected success to clear the previous failure reason');
TcUnit.TEST_FINISHED();
END_METHOD

(* transferTo moves records to another queue without copying them and keeps their FIFO order, so a batch can be handed on without new allocations. *)
METHOD testTransfersQueueOwnership : REFERENCE TO FB_Test
VAR
	source: FB_LogRecordQueue(maxCount:=2);
	destination: FB_LogRecordQueue(maxCount:=2);
	pRecord: POINTER TO FB_LogRecord;
	pFirstOriginal: POINTER TO FB_LogRecord;
	pSecondOriginal: POINTER TO FB_LogRecord;
	failureReason: E_LogRecordQueueFailureReason;
	noFailure: E_LogRecordQueueFailureReason;
	success: BOOL;
	_idx: UDINT;
END_VAR
TcUnit.TEST('testTransfersQueueOwnership');
	noFailure := E_LogRecordQueueFailureReason.NA;
	FOR _idx := 1 TO 2 DO
		// opaque queue node: no factory hands a test an owned FB_LogRecord
		pRecord := __NEW(FB_LogRecord(severityNumber:=E_SeverityNumber.INFO, timestamp:=_idx));
		IF _idx = 1 THEN
			pFirstOriginal := pRecord;
		ELSE
			pSecondOriginal := pRecord;
		END_IF
		success := source.push(pValue:=pRecord, failureReason=>failureReason);
		THIS^.AssertTrue(success, 'Expected source push to succeed');
	END_FOR

	success := source.transferTo(destination:=destination, count:=2, failureReason=>failureReason);
	THIS^.AssertTrue(success AND_THEN failureReason = noFailure, 'Expected queue ownership transfer to succeed');
	THIS^.AssertTrue(source.count = 0 AND_THEN destination.count = 2, 'Expected only the destination to own the records');

	success := destination.pop(pValue:=pRecord, failureReason=>failureReason);
	THIS^.AssertTrue(success AND_THEN pRecord = pFirstOriginal AND_THEN pRecord^.timestamp = 1, 'Expected transfer to preserve the first allocation and FIFO order');
	IF pRecord <> 0 THEN pRecord^.delete(pSelf:=pRecord); END_IF
	success := destination.pop(pValue:=pRecord, failureReason=>failureReason);
	THIS^.AssertTrue(success AND_THEN pRecord = pSecondOriginal AND_THEN pRecord^.timestamp = 2, 'Expected destination to own the same tail allocation');
	IF pRecord <> 0 THEN pRecord^.delete(pSelf:=pRecord); END_IF
TcUnit.TEST_FINISHED();
END_METHOD

(* transferTo moves only the requested number of oldest records and leaves the rest in the source, so a processor can export part of its queue. *)
METHOD testTransfersRequestedCount : REFERENCE TO FB_Test
VAR
	source: FB_LogRecordQueue(maxCount:=3);
	destination: FB_LogRecordQueue(maxCount:=0);
	pRecord: POINTER TO FB_LogRecord;
	failureReason: E_LogRecordQueueFailureReason;
	noFailure: E_LogRecordQueueFailureReason;
	success: BOOL;
	_idx: UDINT;
END_VAR
TcUnit.TEST('testTransfersRequestedCount');
	noFailure := E_LogRecordQueueFailureReason.NA;
	FOR _idx := 1 TO 3 DO
		// opaque queue node: no factory hands a test an owned FB_LogRecord
		pRecord := __NEW(FB_LogRecord(severityNumber:=E_SeverityNumber.INFO, timestamp:=_idx));
		success := source.push(pValue:=pRecord, failureReason=>failureReason);
		THIS^.AssertTrue(success, 'Expected source push to succeed');
	END_FOR

	success := source.transferTo(destination:=destination, count:=2, failureReason=>failureReason);
	THIS^.AssertTrue(success AND_THEN failureReason = noFailure, 'Expected a partial queue transfer to succeed');
	THIS^.AssertTrue(source.count = 1 AND_THEN destination.count = 2, 'Expected the destination to take only the requested count');

	success := destination.pop(pValue:=pRecord, failureReason=>failureReason);
	THIS^.AssertTrue(success AND_THEN pRecord <> 0 AND_THEN pRecord^.timestamp = 1, 'Expected the destination to receive the oldest record first');
	IF pRecord <> 0 THEN pRecord^.delete(pSelf:=pRecord); END_IF
	success := destination.pop(pValue:=pRecord, failureReason=>failureReason);
	THIS^.AssertTrue(success AND_THEN pRecord <> 0 AND_THEN pRecord^.timestamp = 2, 'Expected the destination to receive a FIFO slice');
	IF pRecord <> 0 THEN pRecord^.delete(pSelf:=pRecord); END_IF
	success := source.pop(pValue:=pRecord, failureReason=>failureReason);
	THIS^.AssertTrue(success AND_THEN pRecord <> 0 AND_THEN pRecord^.timestamp = 3, 'Expected the source to retain the untransferred tail');
	IF pRecord <> 0 THEN pRecord^.delete(pSelf:=pRecord); END_IF
TcUnit.TEST_FINISHED();
END_METHOD

END_FUNCTION_BLOCK

// ---- TEST/LOGGING/LOGGER/FB_TestLogger.TcPOU
(* Tests the public logger API. *)
FUNCTION_BLOCK FB_TestLogger EXTENDS FB_TestSuite

THIS^.testEmitWithoutRecordReturnsFailure();
THIS^.testEmitReturnsFirstFluentFailure();
THIS^.testStartingSecondRecordReturnsFailure();
THIS^.testStartLogRecordStampsUnixEpochNanos();
THIS^.testSetTraceContextFromSpanCopiesIdsAndFlags();
THIS^.testSetTraceContextFromSpanWithoutSpanIsNoOp();
THIS^.testSetFlagsStoresTraceFlags();
THIS^.testExitReleasesRecordUnlessCopied();

(*
	When several fluent setters fail, emit reports the first failure and frees the
	incomplete record, so the caller sees the root cause and nothing leaks.
*)
METHOD testEmitReturnsFirstFluentFailure : REFERENCE TO FB_Test
VAR
	resource: FB_Resource('');
	provider: FB_LoggerProvider(resource);
	scope: FB_InstrumentationScope('name', 'version', '');
	logger: FB_Logger(scope, provider);
	success: BOOL;
	failureResult: E_LoggerFailureReason;
END_VAR
TcUnit.TEST('testEmitReturnsFirstFluentFailure');
	// both setters get a deliberately null pointer; the span ID failure comes first
	logger
		.startLogRecord(E_SeverityNumber.ERROR)
		._setSpanId(pBytes:=0, nSize:=0)
		._setTraceId(pBytes:=0, nSize:=0);

	success := logger.emit(failureResult=>failureResult);
	THIS^.AssertFalse(success, 'Expected the invalid Span ID to fail emission');
	THIS^.AssertTrue(
		failureResult = E_LoggerFailureReason.SPAN_ID_BYTES_POINTER_NULL,
		'Expected emit to report the first fluent failure, SPAN_ID_BYTES_POINTER_NULL'
	);
	THIS^.AssertTrue(logger.pLogRecord = 0, 'Expected failed emit to release the incomplete record');
TcUnit.TEST_FINISHED();
END_METHOD

(*
	Calling emit with no record started fails with LOG_RECORD_NOT_STARTED, so a
	misordered call is reported instead of emitting an empty record.
*)
METHOD testEmitWithoutRecordReturnsFailure : REFERENCE TO FB_Test
VAR
	resource: FB_Resource('');
	provider: FB_LoggerProvider(resource);
	scope: FB_InstrumentationScope('name', 'version', '');
	logger: FB_Logger(scope, provider);
	success: BOOL;
	failureResult: E_LoggerFailureReason;
END_VAR
TcUnit.TEST('testEmitWithoutRecordReturnsFailure');
	logger.reset();
	success := logger.emit(failureResult=>failureResult);
	THIS^.AssertFalse(success, 'Expected emit without a started record to fail');
	THIS^.AssertTrue(
		failureResult = E_LoggerFailureReason.LOG_RECORD_NOT_STARTED,
		'Expected emit without a started record to report LOG_RECORD_NOT_STARTED'
	);
TcUnit.TEST_FINISHED();
END_METHOD

(*
	FB_Exit releases a record still being built, so a logger removed mid-chain does not leak it.
	During an online change the copied instance keeps the record, so FB_Exit leaves it alone.
*)
METHOD testExitReleasesRecordUnlessCopied : REFERENCE TO FB_Test
VAR
	resource: FB_Resource('');
	provider: FB_LoggerProvider(resource);
	scope: FB_InstrumentationScope('name', 'version', '');
	logger: FB_Logger(scope, provider);
END_VAR
TcUnit.TEST('testExitReleasesRecordUnlessCopied');
	logger.startLogRecord(E_SeverityNumber.INFO);
	THIS^.AssertTrue(logger.pLogRecord <> 0, 'Expected the logger to hold the record');

	logger.FB_Exit(bInCopyCode:=TRUE);
	THIS^.AssertTrue(logger.pLogRecord <> 0, 'Expected an online change to keep the record');

	logger.FB_Exit(bInCopyCode:=FALSE);
	THIS^.AssertTrue(logger.pLogRecord = 0, 'Expected FB_Exit to release the record');
TcUnit.TEST_FINISHED();
END_METHOD

(*
	_setFlags stores the W3C trace flags in the record's flags, and a later call replaces them.
	The serializer, not the record, leaves flags out for a record without a trace id.
*)
METHOD testSetFlagsStoresTraceFlags : REFERENCE TO FB_Test
VAR
	resource: FB_Resource('');
	provider: FB_LoggerProvider(resource);
	scope: FB_InstrumentationScope('name', 'version', '');
	logger: FB_Logger(scope, provider);
	success: BOOL;
	failureResult: E_LoggerFailureReason;
END_VAR
TcUnit.TEST('testSetFlagsStoresTraceFlags');
	logger
		.startLogRecord(E_SeverityNumber.INFO)
		._setFlags(16#FF);
	THIS^.AssertTrue(logger.pLogRecord <> 0, 'Expected the logger to hold the record');
	IF logger.pLogRecord <> 0 THEN
		THIS^.AssertEquals_UDINT(16#FF, logger.pLogRecord^.flags, 'Expected _setFlags to store all eight trace flag bits');
	END_IF

	logger._setFlags(16#01);  // sampled
	IF logger.pLogRecord <> 0 THEN
		THIS^.AssertEquals_UDINT(1, logger.pLogRecord^.flags, 'Expected a later _setFlags to replace the trace flags');
	END_IF

	success := logger.emit(failureResult=>failureResult);
	THIS^.AssertTrue(success, 'Expected the record to be emitted');
	provider.tick();
TcUnit.TEST_FINISHED();
END_METHOD

(*
	setTraceContextFromSpan copies the span's trace id, span id and W3C trace flags onto the record, so a log
	correlates with its span and is marked sampled only when the span is.
*)
METHOD testSetTraceContextFromSpanCopiesIdsAndFlags : REFERENCE TO FB_Test
VAR
	resource: FB_Resource('');
	loggerProvider: FB_LoggerProvider(resource);
	scope: FB_InstrumentationScope('name', 'version', '');
	logger: FB_Logger(scope, loggerProvider);
	idGenerator: FB_MockIdGenerator;
	tracerProvider: FB_TracerProvider(resource:=resource, idGenerator:=idGenerator, sampler:=TcOtlp_GVL.defaultSampler);
	tracer: FB_Tracer(scope:=scope, provider:=tracerProvider);
	unsampled: STRING(55) := '00-4bf92f3577b34da6a3ce929d0e0e4736-00f067aa0ba902b7-00';
	pUnsampledParent: POINTER TO FB_SpanContext;
	pSampledSpan: POINTER TO FB_Span;
	pUnsampledSpan: POINTER TO FB_Span;
	success: BOOL;
	failureResult: E_LoggerFailureReason;
END_VAR
TcUnit.TEST('testSetTraceContextFromSpanCopiesIdsAndFlags');
	// the default sampler samples a root span and keeps the child of an unsampled parent unsampled
	TraceContextPropagator.extract(pDest:=pUnsampledParent, traceparent:=unsampled, tracestate:='');
	tracer.startSpan(name:='sampled').build(pDest:=pSampledSpan);
	tracer.startSpan(name:='unsampled').setParentUsingContext(pContext:=pUnsampledParent).build(pDest:=pUnsampledSpan);
	THIS^.AssertTrue(pSampledSpan <> 0 AND pUnsampledSpan <> 0, 'Expected both spans to be built');

	IF pSampledSpan <> 0 THEN
		logger
			.startLogRecord(E_SeverityNumber.INFO)
			.setTraceContextFromSpan(pSampledSpan);
		THIS^.AssertTrue(logger.pLogRecord <> 0, 'Expected the logger to hold the record from the sampled span');
		IF logger.pLogRecord <> 0 THEN
			THIS^.AssertTrue(
				logger.pLogRecord^.traceId <> 0 AND_THEN logger.pLogRecord^.traceId <> pSampledSpan^.traceId
				AND_THEN MEMCMP(ADR(logger.pLogRecord^.traceId^.bytes), ADR(pSampledSpan^.traceId^.bytes), SIZEOF(pSampledSpan^.traceId^.bytes)) = 0,
				'Expected the record to own a copy of the span trace id'
			);
			THIS^.AssertTrue(
				logger.pLogRecord^.spanId <> 0 AND_THEN logger.pLogRecord^.spanId <> pSampledSpan^.spanId
				AND_THEN MEMCMP(ADR(logger.pLogRecord^.spanId^.bytes), ADR(pSampledSpan^.spanId^.bytes), SIZEOF(pSampledSpan^.spanId^.bytes)) = 0,
				'Expected the record to own a copy of the span id'
			);
			THIS^.AssertEquals_UDINT(1, logger.pLogRecord^.flags, 'Expected a record from a sampled span to carry the sampled flag');
		END_IF
		success := logger.emit(failureResult=>failureResult);
		THIS^.AssertTrue(success, 'Expected the record from the sampled span to be emitted');
	END_IF

	IF pUnsampledSpan <> 0 THEN
		logger
			.startLogRecord(E_SeverityNumber.INFO)
			.setTraceContextFromSpan(pUnsampledSpan);
		THIS^.AssertTrue(logger.pLogRecord <> 0, 'Expected the logger to hold the record from the unsampled span');
		IF logger.pLogRecord <> 0 THEN
			THIS^.AssertTrue(logger.pLogRecord^.traceId <> 0, 'Expected a record from an unsampled span to keep its trace id');
			THIS^.AssertEquals_UDINT(0, logger.pLogRecord^.flags, 'Expected a record from an unsampled span not to carry the sampled flag');
		END_IF
		success := logger.emit(failureResult=>failureResult);
		THIS^.AssertTrue(success, 'Expected the record from the unsampled span to be emitted');
	END_IF

	loggerProvider.tick();
	IF pSampledSpan <> 0 THEN pSampledSpan^.delete(pSelf:=pSampledSpan); END_IF
	IF pUnsampledSpan <> 0 THEN pUnsampledSpan^.delete(pSelf:=pUnsampledSpan); END_IF
	IF pUnsampledParent <> 0 THEN pUnsampledParent^.delete(pSelf:=pUnsampledParent); END_IF
TcUnit.TEST_FINISHED();
END_METHOD

(*
	setTraceContextFromSpan with a null span, or a span that has no ids, leaves the record without ids and does
	not fail the chain, so the same logging code works inside and outside a span.
*)
METHOD testSetTraceContextFromSpanWithoutSpanIsNoOp : REFERENCE TO FB_Test
VAR
	resource: FB_Resource('');
	provider: FB_LoggerProvider(resource);
	scope: FB_InstrumentationScope('name', 'version', '');
	logger: FB_Logger(scope, provider);
	spanWithoutIds: FB_Span;  // declared directly because the tracer never builds a span without ids
	success: BOOL;
	failureResult: E_LoggerFailureReason;
END_VAR
TcUnit.TEST('testSetTraceContextFromSpanWithoutSpanIsNoOp');
	logger
		.startLogRecord(E_SeverityNumber.INFO)
		.setTraceContextFromSpan(0);
	THIS^.AssertTrue(logger.pLogRecord <> 0, 'Expected the logger to hold the record after a null span');
	IF logger.pLogRecord <> 0 THEN
		THIS^.AssertTrue(logger.pLogRecord^.traceId = 0 AND logger.pLogRecord^.spanId = 0, 'Expected a null span to leave the record without ids');
	END_IF
	success := logger.emit(failureResult=>failureResult);
	THIS^.AssertTrue(success, 'Expected a null span not to fail emission');

	logger
		.startLogRecord(E_SeverityNumber.INFO)
		.setTraceContextFromSpan(ADR(spanWithoutIds));
	THIS^.AssertTrue(logger.pLogRecord <> 0, 'Expected the logger to hold the record after a span without ids');
	IF logger.pLogRecord <> 0 THEN
		THIS^.AssertTrue(logger.pLogRecord^.traceId = 0 AND logger.pLogRecord^.spanId = 0, 'Expected a span without ids to leave the record without ids');
	END_IF
	success := logger.emit(failureResult=>failureResult);
	THIS^.AssertTrue(success, 'Expected a span without ids not to fail emission');

	provider.tick();
TcUnit.TEST_FINISHED();
END_METHOD

(*
	Starting a second record before the first is emitted fails the pending emit and
	frees the record, so one logger never holds or leaks two records at once.
*)
METHOD testStartingSecondRecordReturnsFailure : REFERENCE TO FB_Test
VAR
	resource: FB_Resource('');
	provider: FB_LoggerProvider(resource);
	scope: FB_InstrumentationScope('name', 'version', '');
	logger: FB_Logger(scope, provider);
	success: BOOL;
	failureResult: E_LoggerFailureReason;
END_VAR
TcUnit.TEST('testStartingSecondRecordReturnsFailure');
	logger.startLogRecord(E_SeverityNumber.INFO);
	// deliberately start a second record before the first is emitted
	logger.startLogRecord(E_SeverityNumber.WARN);

	success := logger.emit(failureResult=>failureResult);
	THIS^.AssertFalse(success, 'Expected starting a second record to fail emission');
	THIS^.AssertTrue(
		failureResult = E_LoggerFailureReason.LOG_RECORD_ALREADY_STARTED,
		'Expected starting a second record to report LOG_RECORD_ALREADY_STARTED'
	);
	THIS^.AssertTrue(logger.pLogRecord = 0, 'Expected failed emit to release the incomplete record');
TcUnit.TEST_FINISHED();
END_METHOD

(*
	The auto-stamped timestamp is nanoseconds since the unix epoch. A precedence
	error in (F_GetSystemTime() - DIFF * 100) once underflowed ULINT and produced
	timestamps billions of years in the future.
*)
METHOD testStartLogRecordStampsUnixEpochNanos : REFERENCE TO FB_Test
VAR
	resource: FB_Resource('');
	provider: FB_LoggerProvider(resource);
	scope: FB_InstrumentationScope('name', 'version', '');
	logger: FB_Logger(scope, provider);
	success: BOOL;
	failureResult: E_LoggerFailureReason;
	beforeNs: ULINT;
	afterNs: ULINT;
END_VAR
VAR CONSTANT
	UNIX_EPOCH_DIFF: ULINT := 116444736000000000;  // 1601 -> 1970 offset in 100ns intervals
END_VAR
TcUnit.TEST('testStartLogRecordStampsUnixEpochNanos');
	beforeNs := (F_GetSystemTime() - UNIX_EPOCH_DIFF) * 100;
	logger.startLogRecord(E_SeverityNumber.INFO);
	afterNs := (F_GetSystemTime() - UNIX_EPOCH_DIFF) * 100;

	THIS^.AssertTrue(logger.pLogRecord <> 0, 'Expected startLogRecord to allocate a record');
	IF logger.pLogRecord <> 0 THEN
		THIS^.AssertTrue(
			logger.pLogRecord^.timestamp >= beforeNs AND_THEN logger.pLogRecord^.timestamp <= afterNs,
			'Expected the auto-stamped timestamp to fall within the sampled wall clock window'
		);
	END_IF

	success := logger.emit(failureResult=>failureResult);
	THIS^.AssertTrue(success AND_THEN logger.pLogRecord = 0, 'Expected emit to succeed and release the record');
TcUnit.TEST_FINISHED();
END_METHOD

END_FUNCTION_BLOCK

// ---- TEST/TRACING/TRACER/FB_MockIdGenerator.TcPOU
(* Deterministic id generator for tests. Every identifier is filled with one counter byte,
   so no two identifiers in a test are equal and none is all zero. Set available to FALSE to
   simulate a generator that has nothing ready. *)
FUNCTION_BLOCK FB_MockIdGenerator EXTENDS FB_IdGenerator_Base
VAR_INPUT
	available: BOOL := TRUE;
END_VAR
VAR
	_counter: BYTE;
END_VAR

METHOD generateSpanId : BOOL
VAR_IN_OUT
	spanId: FB_SpanId;
END_VAR
VAR_OUTPUT
	failureReason: E_IdGenFailureReason;
END_VAR
VAR
	_bytes: ARRAY [0..7] OF BYTE;
END_VAR
generateSpanId := FALSE;
failureReason := E_IdGenFailureReason.NA;

IF NOT THIS^.available THEN
	failureReason := E_IdGenFailureReason.NO_IDENTIFIERS_AVAILABLE;
	RETURN;
END_IF

_counter := (_counter MOD 255) + 1;
MEMSET(ADR(_bytes), _counter, SIZEOF(_bytes));
MEMCPY(ADR(spanId.bytes), ADR(_bytes), SIZEOF(spanId.bytes));
generateSpanId := TRUE;
END_METHOD

METHOD generateTraceId : BOOL
VAR_IN_OUT
	traceId: FB_TraceId;
END_VAR
VAR_OUTPUT
	failureReason: E_IdGenFailureReason;
END_VAR
VAR
	_bytes: ARRAY [0..15] OF BYTE;
END_VAR
generateTraceId := FALSE;
failureReason := E_IdGenFailureReason.NA;

IF NOT THIS^.available THEN
	failureReason := E_IdGenFailureReason.NO_IDENTIFIERS_AVAILABLE;
	RETURN;
END_IF

_counter := (_counter MOD 255) + 1;
MEMSET(ADR(_bytes), _counter, SIZEOF(_bytes));
MEMCPY(ADR(traceId.bytes), ADR(_bytes), SIZEOF(traceId.bytes));
generateTraceId := TRUE;
END_METHOD

METHOD tick : BOOL
VAR_OUTPUT
	failureReason: E_IdGenFailureReason;
END_VAR
tick := TRUE;
failureReason := E_IdGenFailureReason.NA;
END_METHOD

END_FUNCTION_BLOCK

// ---- TEST/LOGGING/PROVIDER/FB_TestLoggerProvider.TcPOU
(* Tests FB_LoggerProvider processor registration. *)
FUNCTION_BLOCK FB_TestLoggerProvider EXTENDS FB_TestSuite

THIS^.testStageProcessorChaining();
THIS^.testStageProcessorCount();
THIS^.testTickUnstagesProcessors();
THIS^.testDuplicateProcessorReceivesRecordOnce();
THIS^.testDistinctProcessorsEachReceiveRecord();
THIS^.testTickReportsSuccess();

(*
	Two distinct processors registered with the same provider should each
	receive the emitted record independently.
*)
METHOD testDistinctProcessorsEachReceiveRecord : REFERENCE TO FB_Test
VAR
	resource: FB_Resource('');
	provider: FB_LoggerProvider(resource);
	scope: FB_InstrumentationScope('scope', '1.0.0', '');
	logger: FB_Logger(scope, provider);
	exporterA: FB_LogRecordExporter_ForInspection;
	processorA: FB_LogRecordProcessor_Simple(exporterA);
	exporterB: FB_LogRecordExporter_ForInspection;
	processorB: FB_LogRecordProcessor_Simple(exporterB);
END_VAR
TcUnit.TEST('testDistinctProcessorsEachReceiveRecord');
	provider.stageProcessor(processorA);
	provider.stageProcessor(processorB);

	logger.startLogRecord(severityNumber:=E_SeverityNumber.INFO).emit();
	provider.tick();

	THIS^.AssertEquals_UDINT(1, exporterA.records.count, 'Expected one record in exporter A');
	THIS^.AssertEquals_UDINT(1, exporterB.records.count, 'Expected one record in exporter B');
TcUnit.TEST_FINISHED();
END_METHOD

(*
	When the same processor is added twice (duplicate rejected), it should
	receive each emitted record exactly once — not twice.
*)
METHOD testDuplicateProcessorReceivesRecordOnce : REFERENCE TO FB_Test
VAR
	resource: FB_Resource('');
	provider: FB_LoggerProvider(resource);
	scope: FB_InstrumentationScope('scope', '1.0.0', '');
	logger: FB_Logger(scope, provider);
	exporter: FB_LogRecordExporter_ForInspection;
	processor: FB_LogRecordProcessor_Simple(exporter);
END_VAR
TcUnit.TEST('testDuplicateProcessorReceivesRecordOnce');
	provider.stageProcessor(processor);
	// the second stage of the same processor is silently ignored
	provider.stageProcessor(processor);
	THIS^.AssertEquals_UDINT(1, provider.stagedProcessorCount, 'Expected staging the same processor twice to leave one staged processor');

	logger.startLogRecord(severityNumber:=E_SeverityNumber.INFO).emit();
	provider.tick();

	THIS^.AssertEquals_UDINT(1, exporter.records.count, 'Expected exactly one record in exporter, not two');
TcUnit.TEST_FINISHED();
END_METHOD

(*
	Staging lasts one tick: tick releases every staged processor node, so the
	caller must stage processors again each cycle and no list node leaks.
*)
METHOD testTickUnstagesProcessors : REFERENCE TO FB_Test
VAR
	resource: FB_Resource('');
	provider: FB_LoggerProvider(resource);
	processorA: FB_LogRecordProcessor_Simple(0);
	processorB: FB_LogRecordProcessor_Simple(0);
END_VAR
TcUnit.TEST('testTickUnstagesProcessors');
	provider.stageProcessor(processorA);
	provider.stageProcessor(processorB);
	THIS^.AssertEquals_UDINT(2, provider.stagedProcessorCount, 'Expected two staged processors before tick');
	provider.tick();
	THIS^.AssertEquals_UDINT(0, provider.stagedProcessorCount, 'Expected tick to unstage every processor');
TcUnit.TEST_FINISHED();
END_METHOD

(*
	stageProcessor returns the provider, so processors can be staged in one
	fluent chain and each chained call still counts.
*)
METHOD testStageProcessorChaining : REFERENCE TO FB_Test
VAR
	resource: FB_Resource('');
	provider: FB_LoggerProvider(resource);
	processorA: FB_LogRecordProcessor_Simple(0);
	processorB: FB_LogRecordProcessor_Simple(0);
END_VAR
TcUnit.TEST('testStageProcessorChaining');
	provider.stageProcessor(processorA).stageProcessor(processorB);
	THIS^.AssertEquals_UDINT(2, provider.stagedProcessorCount, 'Expected two staged processors after a chained stageProcessor call');
TcUnit.TEST_FINISHED();
END_METHOD

(*
	stagedProcessorCount starts at zero and rises by one per distinct staged
	processor; tick relies on it to bound its walk of the processor list.
*)
METHOD testStageProcessorCount : REFERENCE TO FB_Test
VAR
	resource: FB_Resource('');
	provider: FB_LoggerProvider(resource);
	processorA: FB_LogRecordProcessor_Simple(0);
	processorB: FB_LogRecordProcessor_Simple(0);
END_VAR
TcUnit.TEST('testStageProcessorCount');
	THIS^.AssertEquals_UDINT(0, provider.stagedProcessorCount, 'Expected zero staged processors after init');
	provider.stageProcessor(processorA);
	THIS^.AssertEquals_UDINT(1, provider.stagedProcessorCount, 'Expected one staged processor after the first stageProcessor call');
	provider.stageProcessor(processorB);
	THIS^.AssertEquals_UDINT(2, provider.stagedProcessorCount, 'Expected two staged processors after the second stageProcessor call');
TcUnit.TEST_FINISHED();
END_METHOD

(*
	Exhausting the staged-processor list is normal loop termination, not a
	corrupt list, so tick must report success once every processor has run.
*)
METHOD testTickReportsSuccess : REFERENCE TO FB_Test
VAR
	resource: FB_Resource('');
	provider: FB_LoggerProvider(resource);
	scope: FB_InstrumentationScope('scope', '1.0.0', '');
	logger: FB_Logger(scope, provider);
	exporterA: FB_LogRecordExporter_ForInspection;
	processorA: FB_LogRecordProcessor_Simple(exporterA);
	exporterB: FB_LogRecordExporter_ForInspection;
	processorB: FB_LogRecordProcessor_Simple(exporterB);
	tickSucceeded: BOOL;
	tickFailureReason: E_LoggerProviderFailureReason;
END_VAR
TcUnit.TEST('testTickReportsSuccess');
	// a single staged processor walks the list to its tail on the first iteration
	logger.startLogRecord(severityNumber:=E_SeverityNumber.INFO).emit();
	tickSucceeded := provider
		.stageProcessor(processorA)
		.tick(failureReason=>tickFailureReason);
	THIS^.AssertTrue(tickSucceeded, 'Expected tick to succeed with one staged processor');
	THIS^.AssertEquals_UDINT(
		TO_UDINT(E_LoggerProviderFailureReason.NA),
		TO_UDINT(tickFailureReason),
		'Expected no failure reason with one staged processor'
	);

	// tick unstages every processor, so both must be staged again
	logger.startLogRecord(severityNumber:=E_SeverityNumber.INFO).emit();
	tickSucceeded := provider
		.stageProcessor(processorA)
		.stageProcessor(processorB)
		.tick(failureReason=>tickFailureReason);
	THIS^.AssertTrue(tickSucceeded, 'Expected tick to succeed with two staged processors');
	THIS^.AssertEquals_UDINT(
		TO_UDINT(E_LoggerProviderFailureReason.NA),
		TO_UDINT(tickFailureReason),
		'Expected no failure reason with two staged processors'
	);

	// a tick with nothing staged still reports success
	tickSucceeded := provider.tick(failureReason=>tickFailureReason);
	THIS^.AssertTrue(tickSucceeded, 'Expected tick to succeed with no staged processors');
TcUnit.TEST_FINISHED();
END_METHOD

END_FUNCTION_BLOCK

// ---- TEST/LOGGING/EXPORTING/UTILS/FB_LogRecordExporter_ForInspection.TcPOU
(*
	Exporter test double that captures the linked list a processor transfers via
	export, so tests can assert on the exported batch. Set busy to
	simulate an exporter that cannot accept a batch. callsWhileBusy counts
	export calls made while busy, which a processor must never make.
*)
FUNCTION_BLOCK FB_LogRecordExporter_ForInspection EXTENDS FB_LogRecordExporter_Base
VAR_INPUT
	busy: BOOL;		// TRUE simulates a busy exporter that refuses batches
END_VAR
VAR_OUTPUT
	callsWhileBusy: UDINT;
END_VAR

METHOD isBusy : BOOL
isBusy := THIS^.busy;
END_METHOD

// the captured batch, for test assertions
PROPERTY records : REFERENCE TO FB_LogRecordQueue
GET
records REF= THIS^._records;
END_GET
END_PROPERTY

METHOD tick : BOOL
VAR_OUTPUT
	failureReason: E_LogRecordExporterFailureReason;
END_VAR
failureReason := E_LogRecordExporterFailureReason.NA;
tick := TRUE;
END_METHOD

METHOD export : BOOL
VAR_IN_OUT
	logRecords: FB_LogRecordQueue;
END_VAR
VAR_INPUT
	count: UDINT;
END_VAR
VAR_OUTPUT
	failureReason: E_LogRecordExporterFailureReason;
END_VAR
IF THIS^.isBusy() THEN
	THIS^.callsWhileBusy := THIS^.callsWhileBusy + 1;
END_IF
export := SUPER^.export(logRecords:=logRecords, count:=count, failureReason=>failureReason);
END_METHOD

END_FUNCTION_BLOCK

// ---- TEST/LOGGING/PROCESSOR/FB_TestLogProcessors.TcPOU
(* Tests simple and batch log processors. *)
FUNCTION_BLOCK FB_TestLogProcessors EXTENDS FB_TestSuite

THIS^.testSimpleProcessorExportsEachRecord();
THIS^.testBatchProcessorQueuesAndFlushes();
THIS^.testProcessorsSkipBusyExporter();

(*
	The batch processor queues emitted records in arrival order (oldest at
	the head), dropping the oldest when the queue is full. Flushing moves
	the oldest maxExportBatchSize records into the exporter's queue, on a
	full batch or when the schedule delay elapses, so records leave in order
	and memory stays bounded however fast the PLC logs. queuedCount reports
	the records waiting for export, and droppedCount the records lost.

	FB_LoggerProvider.tick() unstages every processor, so a processor must be
	staged again before each tick.
*)
METHOD testBatchProcessorQueuesAndFlushes : REFERENCE TO FB_Test
VAR
	resourceA: FB_Resource('resource.a');
	resourceB: FB_Resource('resource.b');
	providerA: FB_LoggerProvider(resourceA);
	providerB: FB_LoggerProvider(resourceB);
	scopeA: FB_InstrumentationScope('scope.a', '1.0.0', '');
	scopeB: FB_InstrumentationScope('scope.b', '1.0.0', '');
	loggerAA: FB_Logger(scopeA, providerA);
	loggerAB: FB_Logger(scopeB, providerA);
	loggerBA: FB_Logger(scopeA, providerB);
	exporter: FB_LogRecordExporter_ForInspection;
	processor: FB_LogRecordProcessor_ForBatchInspection(
		maxQueueSize:=10,
		scheduledDelayMillis:=1000,
		maxExportBatchSize:=6,
		exporter:=exporter
	);
	// no exporter, so onEmit only enriches and never queues
	orphanProcessor: FB_LogRecordProcessor_ForBatchInspection(
		maxQueueSize:=10,
		scheduledDelayMillis:=1000,
		maxExportBatchSize:=6,
		exporter:=0
	);
	boundedExporter: FB_LogRecordExporter_ForInspection;
	boundedProcessor: FB_LogRecordProcessor_ForBatchInspection(
		maxQueueSize:=2,
		scheduledDelayMillis:=1000,
		maxExportBatchSize:=3,
		exporter:=boundedExporter
	);
	timerExporter: FB_LogRecordExporter_ForInspection;
	timerProcessor: FB_LogRecordProcessor_ForBatchInspection(
		maxQueueSize:=0,
		scheduledDelayMillis:=0,
		maxExportBatchSize:=3,
		exporter:=timerExporter
	);
	ts1: ULINT := 1;
	ts2: ULINT := 2;
	ts3: ULINT := 3;
	ts4: ULINT := 4;
	ts5: ULINT := 5;
	ts6: ULINT := 6;
	ts7: ULINT := 7;
	ts8: ULINT := 8;
	ts9: ULINT := 9;
	ts10: ULINT := 10;
	ts11: ULINT := 11;
	ts12: ULINT := 12;
	pRec: POINTER TO FB_LogRecord;
END_VAR
TcUnit.TEST('testBatchProcessorQueuesAndFlushes');
	// processor uses maxExportBatchSize 6 so the count-based flush trigger fires without waiting on the timer

	// --- Scenario: records queue in arrival order ---
	// emit interleaved across (resource, scope) pairs
	loggerBA.startLogRecord(severityNumber:=E_SeverityNumber.INFO).setTimestamp(ts1).emit();
	loggerAB.startLogRecord(severityNumber:=E_SeverityNumber.INFO).setTimestamp(ts2).emit();
	loggerAA.startLogRecord(severityNumber:=E_SeverityNumber.INFO).setTimestamp(ts3).emit();
	loggerBA.startLogRecord(severityNumber:=E_SeverityNumber.INFO).setTimestamp(ts4).emit();
	loggerAA.startLogRecord(severityNumber:=E_SeverityNumber.INFO).setTimestamp(ts5).emit();
	// note, it's bad practice to associate processors with multiple providers
	providerA
		.stageProcessor(processor)
		.tick();
	providerB
		.stageProcessor(processor)
		.tick();
	THIS^.AssertTrue(processor.lastOperationSucceeded, 'Expected the last emit to succeed');
	THIS^.AssertEquals_UDINT(5, processor.records.count, 'Expected five queued records');
	THIS^.AssertEquals_UDINT(5, processor.queuedCount, 'Expected queuedCount to report the five queued records');
	THIS^.AssertEquals_UDINT(0, processor.droppedCount, 'Expected droppedCount to be zero before the queue fills');

	// the queue keeps arrival order per provider, oldest at the head
	processor.records.reset();
	pRec := processor.records.next();
	THIS^.AssertTrue(pRec <> 0 AND_THEN pRec^.timestamp = 2, 'Expected queued record 1 to be ts2');
	pRec := processor.records.next();
	THIS^.AssertTrue(pRec <> 0 AND_THEN pRec^.timestamp = 3, 'Expected queued record 2 to be ts3');
	pRec := processor.records.next();
	THIS^.AssertTrue(pRec <> 0 AND_THEN pRec^.timestamp = 5, 'Expected queued record 3 to be ts5');
	pRec := processor.records.next();
	THIS^.AssertTrue(pRec <> 0 AND_THEN pRec^.timestamp = 1, 'Expected queued record 4 to be ts1');
	pRec := processor.records.next();
	THIS^.AssertTrue(pRec <> 0 AND_THEN pRec^.timestamp = 4, 'Expected queued record 5 to be ts4');
	THIS^.AssertTrue(processor.records.next() = 0, 'Expected queue iteration to be exhausted');

	// --- Scenario: a full batch flushes to the exporter in order ---
	// emit one more to reach maxExportBatchSize, triggering a flush
	loggerAB.startLogRecord(severityNumber:=E_SeverityNumber.INFO).setTimestamp(ts6).emit();
	providerA
		.stageProcessor(processor)
		.tick();
	THIS^.AssertEquals_UDINT(0, processor.records.count, 'Expected zero records left after a full batch flush');
	THIS^.AssertEquals_UDINT(0, processor.queuedCount, 'Expected queuedCount to drop to zero once the batch leaves');
	THIS^.AssertEquals_UDINT(6, exporter.records.count, 'Expected six records in the exported batch');

	// exported batch preserves arrival order
	exporter.records.reset();
	pRec := exporter.records.next();
	THIS^.AssertTrue(pRec <> 0 AND_THEN pRec^.timestamp = 2, 'Expected batch record 0 to be ts2');
	pRec := exporter.records.next();
	THIS^.AssertTrue(pRec <> 0 AND_THEN pRec^.timestamp = 3, 'Expected batch record 1 to be ts3');
	pRec := exporter.records.next();
	THIS^.AssertTrue(pRec <> 0 AND_THEN pRec^.timestamp = 5, 'Expected batch record 2 to be ts5');
	pRec := exporter.records.next();
	THIS^.AssertTrue(pRec <> 0 AND_THEN pRec^.timestamp = 1, 'Expected batch record 3 to be ts1');
	pRec := exporter.records.next();
	THIS^.AssertTrue(pRec <> 0 AND_THEN pRec^.timestamp = 4, 'Expected batch record 4 to be ts4');
	pRec := exporter.records.next();
	THIS^.AssertTrue(pRec <> 0 AND_THEN pRec^.timestamp = 6, 'Expected batch record 5 to be ts6');
	THIS^.AssertTrue(exporter.records.next() = 0, 'Expected batch iteration to be exhausted');

	// --- Scenario: a busy exporter holds records in the queue ---
	// the processor still queues records, but no batch leaves
	exporter.busy := TRUE;
	loggerAB.startLogRecord(severityNumber:=E_SeverityNumber.INFO).setTimestamp(ts7).emit();
	providerA
		.stageProcessor(processor)
		.tick();
	THIS^.AssertEquals_UDINT(1, processor.records.count, 'Expected one queued record while the exporter is busy');
	THIS^.AssertEquals_UDINT(6, exporter.records.count, 'Expected the busy exporter to keep the previous batch');

	// --- Scenario: a partial batch waits for the schedule delay ---
	// once free again, the single queued record stays until scheduledDelayMillis (1000 ms) elapses
	exporter.busy := FALSE;
	providerA
		.stageProcessor(processor)
		.tick();
	THIS^.AssertEquals_UDINT(1, processor.records.count, 'Expected the partial batch to wait for the schedule delay');
	THIS^.AssertEquals_UDINT(6, exporter.records.count, 'Expected no new batch before the schedule delay elapses');

	// --- Scenario: no exporter, no queue ---
	// without a bound exporter onEmit only enriches, so nothing is cloned or queued
	loggerAA.startLogRecord(severityNumber:=E_SeverityNumber.INFO).setTimestamp(ts8).emit();
	providerA
		.stageProcessor(orphanProcessor)
		.tick();
	THIS^.AssertEquals_UDINT(0, orphanProcessor.records.count, 'Expected no queued records without a bound exporter');
	THIS^.AssertTrue(orphanProcessor.lastOperationSucceeded, 'Expected onEmit to succeed without a bound exporter');

	// --- Scenario: a full queue drops the oldest record ---
	// boundedProcessor holds 2 records, so the third emit pushes out the first
	THIS^.AssertEquals_UDINT(2, boundedProcessor.records.maxCount, 'Expected the internal queue to be bounded to maxQueueSize');
	loggerAA.startLogRecord(severityNumber:=E_SeverityNumber.INFO).setTimestamp(ts9).emit();
	loggerAB.startLogRecord(severityNumber:=E_SeverityNumber.INFO).setTimestamp(ts10).emit();
	loggerBA.startLogRecord(severityNumber:=E_SeverityNumber.INFO).setTimestamp(ts11).emit();
	providerA
		.stageProcessor(boundedProcessor)
		.tick();
	providerB
		.stageProcessor(boundedProcessor)
		.tick();
	THIS^.AssertEquals_UDINT(2, boundedProcessor.records.count, 'Expected the queue to stay at maxQueueSize');
	THIS^.AssertEquals_UDINT(1, boundedProcessor.records.droppedCount, 'Expected the oldest record to be dropped');
	THIS^.AssertEquals_UDINT(2, boundedProcessor.queuedCount, 'Expected queuedCount to stay at maxQueueSize');
	THIS^.AssertEquals_UDINT(1, boundedProcessor.droppedCount, 'Expected droppedCount to include the evicted record');
	boundedProcessor.records.reset();
	pRec := boundedProcessor.records.next();
	THIS^.AssertTrue(pRec <> 0 AND_THEN pRec^.timestamp = 10, 'Expected ts9 to be dropped and ts10 at the head');
	pRec := boundedProcessor.records.next();
	THIS^.AssertTrue(pRec <> 0 AND_THEN pRec^.timestamp = 11, 'Expected ts11 at the tail');

	// --- Scenario: the schedule timer flushes a partial batch ---
	// timerProcessor has an unbounded queue (maxQueueSize 0) and a 0 ms delay, so one record is enough to flush
	loggerAA.startLogRecord(severityNumber:=E_SeverityNumber.INFO).setTimestamp(ts12).emit();
	providerA
		.stageProcessor(timerProcessor)
		.tick();
	THIS^.AssertEquals_UDINT(0, timerProcessor.records.count, 'Expected the elapsed timer to flush a partial batch');
	THIS^.AssertEquals_UDINT(0, timerProcessor.queuedCount, 'Expected queuedCount to be zero after the timer flush');
	THIS^.AssertEquals_UDINT(1, timerExporter.records.count, 'Expected one record in the timer-triggered batch');
	timerExporter.records.reset();
	pRec := timerExporter.records.next();
	THIS^.AssertTrue(pRec <> 0 AND_THEN pRec^.timestamp = 12, 'Expected the timer-triggered batch record');

	// --- Cleanup: free releases each processor queue ---
	processor.free();
	orphanProcessor.free();
	boundedProcessor.free();
	timerProcessor.free();
	THIS^.AssertTrue(processor.records.count = 0, 'Expected zero records after free');
	THIS^.AssertTrue(orphanProcessor.records.count = 0, 'Expected zero orphan records after free');
	THIS^.AssertTrue(boundedProcessor.records.count = 0, 'Expected zero bounded records after free');
	THIS^.AssertTrue(timerProcessor.records.count = 0, 'Expected zero timer records after free');
TcUnit.TEST_FINISHED();
END_METHOD

(*
	The simple processor hands each emitted record to an idle exporter straight away, as a clone that
	keeps the body, severity and resource snapshot, so the exporter owns a record that outlives the logger's.
*)
METHOD testSimpleProcessorExportsEachRecord : REFERENCE TO FB_Test
VAR
	resource: FB_Resource('');
	provider: FB_LoggerProvider(resource);
	scope: FB_InstrumentationScope('name', 'version', 'schemaUrl');
	logger: FB_Logger(scope, provider);
	exporter: FB_LogRecordExporter_ForInspection;
	processor: FB_LogRecordProcessor_Simple(exporter);
	pRec: POINTER TO FB_LogRecord;
	pBody: POINTER TO FB_String;
END_VAR
TcUnit.TEST('testSimpleProcessorExportsEachRecord');
	resource.attributes.setStringAttribute('plc.name', 'sim.plc');
	logger.startLogRecord(
			severityNumber:=E_SeverityNumber.ERROR
		)
		.setBody('this is a test')
		.emit();
	provider
		.stageProcessor(processor)
		.tick();

	THIS^.AssertEquals_UDINT(1, exporter.records.count, 'Expected the simple processor to export the emitted record');
	exporter.records.reset();
	pRec := exporter.records.next();
	THIS^.AssertTrue(pRec <> 0, 'Expected the exporter to hold the exported record');
	IF pRec <> 0 THEN
		THIS^.AssertTrue(
			pRec^.severityNumber = E_SeverityNumber.ERROR,
			'Expected the exported record to keep its ERROR severity'
		);
		THIS^.AssertTrue(
			pRec^.body <> 0 AND_THEN pRec^.body^.eType = E_ValueType.E_String,
			'Expected the exported record to keep its string body'
		);
		IF pRec^.body <> 0 AND_THEN pRec^.body^.eType = E_ValueType.E_String THEN
			pBody := pRec^.body;
			THIS^.AssertEquals_STRING('this is a test', pBody^.pString^, 'Expected the exported body text');
		END_IF
		THIS^.AssertEquals_UDINT(1, pRec^.resource.attributes.count, 'Expected the exported record to keep the resource attribute');
	END_IF
	exporter.free();
TcUnit.TEST_FINISHED();
END_METHOD

(* Neither processor calls export on a busy exporter, even when the batch processor has a full batch ready. *)
METHOD testProcessorsSkipBusyExporter : REFERENCE TO FB_Test
VAR
	resource: FB_Resource('');
	provider: FB_LoggerProvider(resource);
	scope: FB_InstrumentationScope('scope', '1.0.0', '');
	logger: FB_Logger(scope, provider);
	simpleExporter: FB_LogRecordExporter_ForInspection;
	simpleProcessor: FB_LogRecordProcessor_Simple(simpleExporter);
	batchExporter: FB_LogRecordExporter_ForInspection;
	batchProcessor: FB_LogRecordProcessor_ForBatchInspection(
		maxQueueSize:=10,
		scheduledDelayMillis:=60000,
		maxExportBatchSize:=1,
		exporter:=batchExporter
	);
END_VAR
TcUnit.TEST('testProcessorsSkipBusyExporter');
	simpleExporter.busy := TRUE;
	batchExporter.busy := TRUE;
	logger.startLogRecord(severityNumber:=E_SeverityNumber.INFO).setBody('work').emit();
	provider
		.stageProcessor(simpleProcessor)
		.stageProcessor(batchProcessor)
		.tick();
	THIS^.AssertEquals_UDINT(0, simpleExporter.callsWhileBusy, 'Expected the simple processor not to call a busy exporter');
	THIS^.AssertEquals_UDINT(0, simpleExporter.records.count, 'Expected the busy simple exporter to receive nothing');
	THIS^.AssertEquals_UDINT(0, batchExporter.callsWhileBusy, 'Expected the batch processor not to call a busy exporter');
	THIS^.AssertEquals_UDINT(1, batchProcessor.records.count, 'Expected the full batch to wait in the processor');
	THIS^.AssertEquals_UDINT(1, batchProcessor.queuedCount, 'Expected queuedCount to include the batch held for a busy exporter');
	THIS^.AssertEquals_UDINT(0, batchProcessor.droppedCount, 'Expected a busy exporter not to make the batch processor drop records');

	batchExporter.busy := FALSE;
	provider
		.stageProcessor(batchProcessor)
		.tick();
	THIS^.AssertEquals_UDINT(1, batchExporter.records.count, 'Expected the batch once the exporter is idle');
	THIS^.AssertEquals_UDINT(0, batchProcessor.records.count, 'Expected the processor queue to be empty');
	THIS^.AssertEquals_UDINT(0, batchProcessor.queuedCount, 'Expected queuedCount to be zero once the held batch is exported');
	simpleExporter.free();
	batchExporter.free();
	batchProcessor.free();
TcUnit.TEST_FINISHED();
END_METHOD

END_FUNCTION_BLOCK

